(* Logix 5000 project; controller TFF vendor 1 type 14 code 107 rev 33.11; software revision 33.04; part 12 of 38 *)

        [5,197].Criteria2Value := -1000000.0, [5,197].ActionValue := -1000000.0, [5,198].Criteria1 := -999, [5,198].Criteria1Operator := -999, [5,198].Boolean := -999, [5,198].Criteria2 := -999, [5,198].Criteria2Operator := -999, [5,198].Action := -999, [5,198].Label := -999, [5,198].Criteria1Value := -1000000.0, [5,198].Criteria2Value := -1000000.0, [5,198].ActionValue := -1000000.0, [5,199].Criteria1 := -999, [5,199].Criteria1Operator := -999, [5,199].Boolean := -999, [5,199].Criteria2 := -999, [5,199].Criteria2Operator := -999, [5,199].Action := -999, [5,199].Label := -999, [5,199].Criteria1Value := -1000000.0, [5,199].Criteria2Value := -1000000.0, [5,199].ActionValue := -1000000.0, [5,200].Criteria1 := -999, [5,200].Criteria1Operator := -999, [5,200].Boolean := -999, [5,200].Criteria2 := -999, [5,200].Criteria2Operator := -999, [5,200].Action := -999, [5,200].Label := -999, [5,200].Criteria1Value := -1000000.0, [5,200].Criteria2Value := -1000000.0, [5,200].ActionValue := -1000000.0, [5,201].Criteria1 := -999, [5,201].Criteria1Operator := -999, [5,201].Boolean := -999, [5,201].Criteria2 := -999, [5,201].Criteria2Operator := -999, [5,201].Action := -999, [5,201].Label := -999, [5,201].Criteria1Value := -1000000.0, [5,201].Criteria2Value := -1000000.0, [5,201].ActionValue := -1000000.0, [5,202].Criteria1 := -999, [5,202].Criteria1Operator := -999, [5,202].Boolean := -999, [5,202].Criteria2 := -999, [5,202].Criteria2Operator := -999, [5,202].Action := -999, [5,202].Label := -999, [5,202].Criteria1Value := -1000000.0, [5,202].Criteria2Value := -1000000.0, [5,202].ActionValue := -1000000.0, [5,203].Criteria1 := -999, [5,203].Criteria1Operator := -999, [5,203].Boolean := -999, [5,203].Criteria2 := -999, [5,203].Criteria2Operator := -999, [5,203].Action := -999, [5,203].Label := -999, [5,203].Criteria1Value := -1000000.0,
        [5,203].Criteria2Value := -1000000.0, [5,203].ActionValue := -1000000.0, [5,204].Criteria1 := -999, [5,204].Criteria1Operator := -999, [5,204].Boolean := -999, [5,204].Criteria2 := -999, [5,204].Criteria2Operator := -999, [5,204].Action := -999, [5,204].Label := -999, [5,204].Criteria1Value := -1000000.0, [5,204].Criteria2Value := -1000000.0, [5,204].ActionValue := -1000000.0, [5,205].Criteria1 := -999, [5,205].Criteria1Operator := -999, [5,205].Boolean := -999, [5,205].Criteria2 := -999, [5,205].Criteria2Operator := -999, [5,205].Action := -999, [5,205].Label := -999, [5,205].Criteria1Value := -1000000.0, [5,205].Criteria2Value := -1000000.0, [5,205].ActionValue := -1000000.0, [5,206].Criteria1 := -999, [5,206].Criteria1Operator := -999, [5,206].Boolean := -999, [5,206].Criteria2 := -999, [5,206].Criteria2Operator := -999, [5,206].Action := -999, [5,206].Label := -999, [5,206].Criteria1Value := -1000000.0, [5,206].Criteria2Value := -1000000.0, [5,206].ActionValue := -1000000.0, [5,207].Criteria1 := -999, [5,207].Criteria1Operator := -999, [5,207].Boolean := -999, [5,207].Criteria2 := -999, [5,207].Criteria2Operator := -999, [5,207].Action := -999, [5,207].Label := -999, [5,207].Criteria1Value := -1000000.0, [5,207].Criteria2Value := -1000000.0, [5,207].ActionValue := -1000000.0, [5,208].Criteria1 := -999, [5,208].Criteria1Operator := -999, [5,208].Boolean := -999, [5,208].Criteria2 := -999, [5,208].Criteria2Operator := -999, [5,208].Action := -999, [5,208].Label := -999, [5,208].Criteria1Value := -1000000.0, [5,208].Criteria2Value := -1000000.0, [5,208].ActionValue := -1000000.0, [5,209].Criteria1 := -999, [5,209].Criteria1Operator := -999, [5,209].Boolean := -999, [5,209].Criteria2 := -999, [5,209].Criteria2Operator := -999, [5,209].Action := -999, [5,209].Label := -999, [5,209].Criteria1Value := -1000000.0,
        [5,209].Criteria2Value := -1000000.0, [5,209].ActionValue := -1000000.0, [5,210].Criteria1 := -999, [5,210].Criteria1Operator := -999, [5,210].Boolean := -999, [5,210].Criteria2 := -999, [5,210].Criteria2Operator := -999, [5,210].Action := -999, [5,210].Label := -999, [5,210].Criteria1Value := -1000000.0, [5,210].Criteria2Value := -1000000.0, [5,210].ActionValue := -1000000.0, [5,211].Criteria1 := -999, [5,211].Criteria1Operator := -999, [5,211].Boolean := -999, [5,211].Criteria2 := -999, [5,211].Criteria2Operator := -999, [5,211].Action := -999, [5,211].Label := -999, [5,211].Criteria1Value := -1000000.0, [5,211].Criteria2Value := -1000000.0, [5,211].ActionValue := -1000000.0, [5,212].Criteria1 := -999, [5,212].Criteria1Operator := -999, [5,212].Boolean := -999, [5,212].Criteria2 := -999, [5,212].Criteria2Operator := -999, [5,212].Action := -999, [5,212].Label := -999, [5,212].Criteria1Value := -1000000.0, [5,212].Criteria2Value := -1000000.0, [5,212].ActionValue := -1000000.0, [5,213].Criteria1 := -999, [5,213].Criteria1Operator := -999, [5,213].Boolean := -999, [5,213].Criteria2 := -999, [5,213].Criteria2Operator := -999, [5,213].Action := -999, [5,213].Label := -999, [5,213].Criteria1Value := -1000000.0, [5,213].Criteria2Value := -1000000.0, [5,213].ActionValue := -1000000.0, [5,214].Criteria1 := -999, [5,214].Criteria1Operator := -999, [5,214].Boolean := -999, [5,214].Criteria2 := -999, [5,214].Criteria2Operator := -999, [5,214].Action := -999, [5,214].Label := -999, [5,214].Criteria1Value := -1000000.0, [5,214].Criteria2Value := -1000000.0, [5,214].ActionValue := -1000000.0, [5,215].Criteria1 := -999, [5,215].Criteria1Operator := -999, [5,215].Boolean := -999, [5,215].Criteria2 := -999, [5,215].Criteria2Operator := -999, [5,215].Action := -999, [5,215].Label := -999, [5,215].Criteria1Value := -1000000.0,
        [5,215].Criteria2Value := -1000000.0, [5,215].ActionValue := -1000000.0, [5,216].Criteria1 := -999, [5,216].Criteria1Operator := -999, [5,216].Boolean := -999, [5,216].Criteria2 := -999, [5,216].Criteria2Operator := -999, [5,216].Action := -999, [5,216].Label := -999, [5,216].Criteria1Value := -1000000.0, [5,216].Criteria2Value := -1000000.0, [5,216].ActionValue := -1000000.0, [5,217].Criteria1 := -999, [5,217].Criteria1Operator := -999, [5,217].Boolean := -999, [5,217].Criteria2 := -999, [5,217].Criteria2Operator := -999, [5,217].Action := -999, [5,217].Label := -999, [5,217].Criteria1Value := -1000000.0, [5,217].Criteria2Value := -1000000.0, [5,217].ActionValue := -1000000.0, [5,218].Criteria1 := -999, [5,218].Criteria1Operator := -999, [5,218].Boolean := -999, [5,218].Criteria2 := -999, [5,218].Criteria2Operator := -999, [5,218].Action := -999, [5,218].Label := -999, [5,218].Criteria1Value := -1000000.0, [5,218].Criteria2Value := -1000000.0, [5,218].ActionValue := -1000000.0, [5,219].Criteria1 := -999, [5,219].Criteria1Operator := -999, [5,219].Boolean := -999, [5,219].Criteria2 := -999, [5,219].Criteria2Operator := -999, [5,219].Action := -999, [5,219].Label := -999, [5,219].Criteria1Value := -1000000.0, [5,219].Criteria2Value := -1000000.0, [5,219].ActionValue := -1000000.0, [5,220].Criteria1 := -999, [5,220].Criteria1Operator := -999, [5,220].Boolean := -999, [5,220].Criteria2 := -999, [5,220].Criteria2Operator := -999, [5,220].Action := -999, [5,220].Label := -999, [5,220].Criteria1Value := -1000000.0, [5,220].Criteria2Value := -1000000.0, [5,220].ActionValue := -1000000.0, [5,221].Criteria1 := -999, [5,221].Criteria1Operator := -999, [5,221].Boolean := -999, [5,221].Criteria2 := -999, [5,221].Criteria2Operator := -999, [5,221].Action := -999, [5,221].Label := -999, [5,221].Criteria1Value := -1000000.0,
        [5,221].Criteria2Value := -1000000.0, [5,221].ActionValue := -1000000.0, [5,222].Criteria1 := -999, [5,222].Criteria1Operator := -999, [5,222].Boolean := -999, [5,222].Criteria2 := -999, [5,222].Criteria2Operator := -999, [5,222].Action := -999, [5,222].Label := -999, [5,222].Criteria1Value := -1000000.0, [5,222].Criteria2Value := -1000000.0, [5,222].ActionValue := -1000000.0, [5,223].Criteria1 := -999, [5,223].Criteria1Operator := -999, [5,223].Boolean := -999, [5,223].Criteria2 := -999, [5,223].Criteria2Operator := -999, [5,223].Action := -999, [5,223].Label := -999, [5,223].Criteria1Value := -1000000.0, [5,223].Criteria2Value := -1000000.0, [5,223].ActionValue := -1000000.0, [5,224].Criteria1 := -999, [5,224].Criteria1Operator := -999, [5,224].Boolean := -999, [5,224].Criteria2 := -999, [5,224].Criteria2Operator := -999, [5,224].Action := -999, [5,224].Label := -999, [5,224].Criteria1Value := -1000000.0, [5,224].Criteria2Value := -1000000.0, [5,224].ActionValue := -1000000.0, [5,225].Criteria1 := -999, [5,225].Criteria1Operator := -999, [5,225].Boolean := -999, [5,225].Criteria2 := -999, [5,225].Criteria2Operator := -999, [5,225].Action := -999, [5,225].Label := -999, [5,225].Criteria1Value := -1000000.0, [5,225].Criteria2Value := -1000000.0, [5,225].ActionValue := -1000000.0, [5,226].Criteria1 := -999, [5,226].Criteria1Operator := -999, [5,226].Boolean := -999, [5,226].Criteria2 := -999, [5,226].Criteria2Operator := -999, [5,226].Action := -999, [5,226].Label := -999, [5,226].Criteria1Value := -1000000.0, [5,226].Criteria2Value := -1000000.0, [5,226].ActionValue := -1000000.0, [5,227].Criteria1 := -999, [5,227].Criteria1Operator := -999, [5,227].Boolean := -999, [5,227].Criteria2 := -999, [5,227].Criteria2Operator := -999, [5,227].Action := -999, [5,227].Label := -999, [5,227].Criteria1Value := -1000000.0,
        [5,227].Criteria2Value := -1000000.0, [5,227].ActionValue := -1000000.0, [5,228].Criteria1 := -999, [5,228].Criteria1Operator := -999, [5,228].Boolean := -999, [5,228].Criteria2 := -999, [5,228].Criteria2Operator := -999, [5,228].Action := -999, [5,228].Label := -999, [5,228].Criteria1Value := -1000000.0, [5,228].Criteria2Value := -1000000.0, [5,228].ActionValue := -1000000.0, [5,229].Criteria1 := -999, [5,229].Criteria1Operator := -999, [5,229].Boolean := -999, [5,229].Criteria2 := -999, [5,229].Criteria2Operator := -999, [5,229].Action := -999, [5,229].Label := -999, [5,229].Criteria1Value := -1000000.0, [5,229].Criteria2Value := -1000000.0, [5,229].ActionValue := -1000000.0, [5,230].Criteria1 := -999, [5,230].Criteria1Operator := -999, [5,230].Boolean := -999, [5,230].Criteria2 := -999, [5,230].Criteria2Operator := -999, [5,230].Action := -999, [5,230].Label := -999, [5,230].Criteria1Value := -1000000.0, [5,230].Criteria2Value := -1000000.0, [5,230].ActionValue := -1000000.0, [5,231].Criteria1 := -999, [5,231].Criteria1Operator := -999, [5,231].Boolean := -999, [5,231].Criteria2 := -999, [5,231].Criteria2Operator := -999, [5,231].Action := -999, [5,231].Label := -999, [5,231].Criteria1Value := -1000000.0, [5,231].Criteria2Value := -1000000.0, [5,231].ActionValue := -1000000.0, [5,232].Criteria1 := -999, [5,232].Criteria1Operator := -999, [5,232].Boolean := -999, [5,232].Criteria2 := -999, [5,232].Criteria2Operator := -999, [5,232].Action := -999, [5,232].Label := -999, [5,232].Criteria1Value := -1000000.0, [5,232].Criteria2Value := -1000000.0, [5,232].ActionValue := -1000000.0, [5,233].Criteria1 := -999, [5,233].Criteria1Operator := -999, [5,233].Boolean := -999, [5,233].Criteria2 := -999, [5,233].Criteria2Operator := -999, [5,233].Action := -999, [5,233].Label := -999, [5,233].Criteria1Value := -1000000.0,
        [5,233].Criteria2Value := -1000000.0, [5,233].ActionValue := -1000000.0, [5,234].Criteria1 := -999, [5,234].Criteria1Operator := -999, [5,234].Boolean := -999, [5,234].Criteria2 := -999, [5,234].Criteria2Operator := -999, [5,234].Action := -999, [5,234].Label := -999, [5,234].Criteria1Value := -1000000.0, [5,234].Criteria2Value := -1000000.0, [5,234].ActionValue := -1000000.0, [5,235].Criteria1 := -999, [5,235].Criteria1Operator := -999, [5,235].Boolean := -999, [5,235].Criteria2 := -999, [5,235].Criteria2Operator := -999, [5,235].Action := -999, [5,235].Label := -999, [5,235].Criteria1Value := -1000000.0, [5,235].Criteria2Value := -1000000.0, [5,235].ActionValue := -1000000.0, [5,236].Criteria1 := -999, [5,236].Criteria1Operator := -999, [5,236].Boolean := -999, [5,236].Criteria2 := -999, [5,236].Criteria2Operator := -999, [5,236].Action := -999, [5,236].Label := -999, [5,236].Criteria1Value := -1000000.0, [5,236].Criteria2Value := -1000000.0, [5,236].ActionValue := -1000000.0, [5,237].Criteria1 := -999, [5,237].Criteria1Operator := -999, [5,237].Boolean := -999, [5,237].Criteria2 := -999, [5,237].Criteria2Operator := -999, [5,237].Action := -999, [5,237].Label := -999, [5,237].Criteria1Value := -1000000.0, [5,237].Criteria2Value := -1000000.0, [5,237].ActionValue := -1000000.0, [5,238].Criteria1 := -999, [5,238].Criteria1Operator := -999, [5,238].Boolean := -999, [5,238].Criteria2 := -999, [5,238].Criteria2Operator := -999, [5,238].Action := -999, [5,238].Label := -999, [5,238].Criteria1Value := -1000000.0, [5,238].Criteria2Value := -1000000.0, [5,238].ActionValue := -1000000.0, [5,239].Criteria1 := -999, [5,239].Criteria1Operator := -999, [5,239].Boolean := -999, [5,239].Criteria2 := -999, [5,239].Criteria2Operator := -999, [5,239].Action := -999, [5,239].Label := -999, [5,239].Criteria1Value := -1000000.0,
        [5,239].Criteria2Value := -1000000.0, [5,239].ActionValue := -1000000.0, [5,240].Criteria1 := -999, [5,240].Criteria1Operator := -999, [5,240].Boolean := -999, [5,240].Criteria2 := -999, [5,240].Criteria2Operator := -999, [5,240].Action := -999, [5,240].Label := -999, [5,240].Criteria1Value := -1000000.0, [5,240].Criteria2Value := -1000000.0, [5,240].ActionValue := -1000000.0, [5,241].Criteria1 := -999, [5,241].Criteria1Operator := -999, [5,241].Boolean := -999, [5,241].Criteria2 := -999, [5,241].Criteria2Operator := -999, [5,241].Action := -999, [5,241].Label := -999, [5,241].Criteria1Value := -1000000.0, [5,241].Criteria2Value := -1000000.0, [5,241].ActionValue := -1000000.0, [5,242].Criteria1 := -999, [5,242].Criteria1Operator := -999, [5,242].Boolean := -999, [5,242].Criteria2 := -999, [5,242].Criteria2Operator := -999, [5,242].Action := -999, [5,242].Label := -999, [5,242].Criteria1Value := -1000000.0, [5,242].Criteria2Value := -1000000.0, [5,242].ActionValue := -1000000.0, [5,243].Criteria1 := -999, [5,243].Criteria1Operator := -999, [5,243].Boolean := -999, [5,243].Criteria2 := -999, [5,243].Criteria2Operator := -999, [5,243].Action := -999, [5,243].Label := -999, [5,243].Criteria1Value := -1000000.0, [5,243].Criteria2Value := -1000000.0, [5,243].ActionValue := -1000000.0, [5,244].Criteria1 := -999, [5,244].Criteria1Operator := -999, [5,244].Boolean := -999, [5,244].Criteria2 := -999, [5,244].Criteria2Operator := -999, [5,244].Action := -999, [5,244].Label := -999, [5,244].Criteria1Value := -1000000.0, [5,244].Criteria2Value := -1000000.0, [5,244].ActionValue := -1000000.0, [5,245].Criteria1 := -999, [5,245].Criteria1Operator := -999, [5,245].Boolean := -999, [5,245].Criteria2 := -999, [5,245].Criteria2Operator := -999, [5,245].Action := -999, [5,245].Label := -999, [5,245].Criteria1Value := -1000000.0,
        [5,245].Criteria2Value := -1000000.0, [5,245].ActionValue := -1000000.0, [5,246].Criteria1 := -999, [5,246].Criteria1Operator := -999, [5,246].Boolean := -999, [5,246].Criteria2 := -999, [5,246].Criteria2Operator := -999, [5,246].Action := -999, [5,246].Label := -999, [5,246].Criteria1Value := -1000000.0, [5,246].Criteria2Value := -1000000.0, [5,246].ActionValue := -1000000.0, [5,247].Criteria1 := -999, [5,247].Criteria1Operator := -999, [5,247].Boolean := -999, [5,247].Criteria2 := -999, [5,247].Criteria2Operator := -999, [5,247].Action := -999, [5,247].Label := -999, [5,247].Criteria1Value := -1000000.0, [5,247].Criteria2Value := -1000000.0, [5,247].ActionValue := -1000000.0, [5,248].Criteria1 := -999, [5,248].Criteria1Operator := -999, [5,248].Boolean := -999, [5,248].Criteria2 := -999, [5,248].Criteria2Operator := -999, [5,248].Action := -999, [5,248].Label := -999, [5,248].Criteria1Value := -1000000.0, [5,248].Criteria2Value := -1000000.0, [5,248].ActionValue := -1000000.0, [5,249].Criteria1 := -999, [5,249].Criteria1Operator := -999, [5,249].Boolean := -999, [5,249].Criteria2 := -999, [5,249].Criteria2Operator := -999, [5,249].Action := -999, [5,249].Label := -999, [5,249].Criteria1Value := -1000000.0, [5,249].Criteria2Value := -1000000.0, [5,249].ActionValue := -1000000.0, [5,250].Criteria1 := -999, [5,250].Criteria1Operator := -999, [5,250].Boolean := -999, [5,250].Criteria2 := -999, [5,250].Criteria2Operator := -999, [5,250].Action := -999, [5,250].Label := -999, [5,250].Criteria1Value := -1000000.0, [5,250].Criteria2Value := -1000000.0, [5,250].ActionValue := -1000000.0);   // Operation Table
        [0,0]   // Null Step
        [1,0]   // Null Step
        [2,0]   // Null Step
        [3,0]   // Null Step
        [4,0]   // Null Step
        [5,0]   // Null Step
   Options : Options := (CCP_Report := 1, InletFeed := 1, FeedTank := 1, TransferFlow := 1, TankPH := 1, FiltrateNoInstrum_Dis := 1, FiltrateCondPHUV := 1, FiltrateUltrasonicFlow := 1, SingleUsePH := 1, External_IO := 1, TFF80 := 1);   // Options List
   PCDateTime : DINT[7] := ([0] := 2025, [1] := 10, [2] := 3, [3] := 11, [4] := 41, [5] := 1, [6] := -1);   // Date/Time Array from PC
   PcToPLCHeartBeat : BOOL;   // PC to PLC communication heartbeat Set to 1 by HMI Reset to 0 by plc
   PCV101 : ALIAS FOR AnalogPoint[3];
   PCV101_AO : ALIAS FOR AnalogOutput[3];
   PCV101_Calib : PCV_Calib;   // PCV101 Position Calibration
   PCV101_Control : PCV_Control := (FullOpenResetTimer.PRE := 3000, FullCloseSP := 100.0, FullCloseResetTimer.PRE := 3000, ClosedStatusSP := 95.0);   // PCV101 Control UDT
   PCV101_CVTune : CVTune := (ClosedRaw := 12340.0, OpenRaw := 27508.0, MaxOutput := 100.0, MinTimer.PRE := 5000, MaxTimer.PRE := 5000);
   PCV101_PID : PCV := (PV := 0.032964136, CV := 100.0, OpenRawValue := 27508.0, ClosedRawValue := 12340.0);   // PCV101 PID Management
   PCV101_SIG : ALIAS FOR DigitalPoint[102];
   PCV101Alarm : ALIAS FOR AlarmAnalog[3];
   PCV201 : ALIAS FOR AnalogPoint[4];
   PCV201_AO : ALIAS FOR AnalogOutput[4];
   PCV201_Calib : PCV_Calib;   // PCV201 Position Calibration
   PCV201_Control : PCV_Control := (FullOpenSP := 100.0, FullOpenResetTimer.PRE := 3000, FullCloseResetTimer.PRE := 3000, ClosedStatusSP := 95.0);   // PCV201 Control UDT
   PCV201_CVTune : CVTune := (ClosedRaw := 25520.0, OpenRaw := 10318.0, MaxOutput := 100.0, MinTimer.PRE := 5000, MaxTimer.PRE := 5000);
   PCV201_PID : PCV := (PV := 51.769505, OpenRawValue := 10318.0, ClosedRawValue := 25520.0);   // PCV201 PID Management
   PCV201_SIG : ALIAS FOR DigitalPoint[103];
   PCV201Alarm : ALIAS FOR AlarmAnalog[4];
   PERM : ALIAS FOR AnalogPoint[46];
   PERMAlarm : ALIAS FOR AlarmAnalog[46];
   Phase : Phases[6] := ([0].Stop := 1, [0].Hold := 1, [0].JumpStep := 13, [0].StartStep := 1, [0].TotalSteps := 16, [0].ActualStep := 12, [1].JumpStep := 51, [1].StartStep := 1, [1].TotalSteps := 49, [1].ActualStep := 50, [2].JumpStep := 11, [2].StartStep := 1, [2].TotalSteps := 9, [2].ActualStep := 10, [3].JumpStep := 14, [3].StartStep := 1, [3].TotalSteps := 45, [3].ActualStep := 13, [4].JumpStep := 68, [4].StartStep := 1, [4].TotalSteps := 66, [4].ActualStep := 67, [5].JumpStep := 6, [5].StartStep := 1, [5].Crit1MetTime := 1, [5].ActualStep := 5);   // Phase Control Array
   Phase0 : ALIAS FOR Phase[0];   // Phase 0
   Phase0_PauseTime : ALIAS FOR Timers[12];   // Phase 0 Pause Time
   Phase0_StepTime : ALIAS FOR Timers[6];   // Phase 0 Step Time
   Phase0_Totalizer_Feed : ALIAS FOR PhaseTotalizer[0];   // Phase 0 Total Feed
   Phase0_Totalizer_Filtrate : ALIAS FOR PhaseTotalizer[6];   // Phase 0 Total Filtrate
   Phase0_Totalizer_Transfer : ALIAS FOR PhaseTotalizer[12];   // Phase 0 Total Transfer
   Phase0_TotalTime : ALIAS FOR Timers[0];   // Phase 0 Total Time
   Phase1 : ALIAS FOR Phase[1];   // Phase 1
   Phase1_PauseTime : ALIAS FOR Timers[13];   // Phase 1 Pause Time
   Phase1_StepTime : ALIAS FOR Timers[7];   // Phase 1 Step Time
   Phase1_Totalizer_Feed : ALIAS FOR PhaseTotalizer[1];   // Phase 1 Total Feed
   Phase1_Totalizer_Filtrate : ALIAS FOR PhaseTotalizer[7];   // Phase 1 Total Filtrate
   Phase1_Totalizer_Transfer : ALIAS FOR PhaseTotalizer[13];   // Phase 1 Total Transfer
   Phase1_TotalTime : ALIAS FOR Timers[1];   // Phase 1 Total Time
   Phase2 : ALIAS FOR Phase[2];   // Phase 2
   Phase2_PauseTime : ALIAS FOR Timers[14];   // Phase 2 Pause Time
   Phase2_StepTime : ALIAS FOR Timers[8];   // Phase 2 Step Time
   Phase2_Totalizer_Feed : ALIAS FOR PhaseTotalizer[2];   // Phase 2 Total Feed
   Phase2_Totalizer_Filtrate : ALIAS FOR PhaseTotalizer[8];   // Phase 2 Total Filtrate
   Phase2_Totalizer_Transfer : ALIAS FOR PhaseTotalizer[14];   // Phase 2 Total Transfer
   Phase2_TotalTime : ALIAS FOR Timers[2];   // Phase 2 Total Time
   Phase3 : ALIAS FOR Phase[3];   // Phase 3
   Phase3_PauseTime : ALIAS FOR Timers[15];   // Phase 3 Pause Time
   Phase3_StepTime : ALIAS FOR Timers[9];   // Phase 3 Step Time
   Phase3_Totalizer_Feed : ALIAS FOR PhaseTotalizer[3];   // Phase 3 Total Feed
   Phase3_Totalizer_Filtrate : ALIAS FOR PhaseTotalizer[9];   // Phase 3 Total Filtrate
   Phase3_Totalizer_Transfer : ALIAS FOR PhaseTotalizer[15];   // Phase 3 Total Transfer
   Phase3_TotalTime : ALIAS FOR Timers[3];   // Phase 3 Total Time
   Phase4 : ALIAS FOR Phase[4];   // Phase 4
   Phase4_PauseTime : ALIAS FOR Timers[16];   // Phase 4 Pause Time
   Phase4_StepTime : ALIAS FOR Timers[10];   // Phase 4 Step Time
   Phase4_Totalizer_Feed : ALIAS FOR PhaseTotalizer[4];   // Phase 4 Total Feed
   Phase4_Totalizer_Filtrate : ALIAS FOR PhaseTotalizer[10];   // Phase 4 Total Filtrate
   Phase4_Totalizer_Transfer : ALIAS FOR PhaseTotalizer[16];   // Phase 4 Total Transfer
   Phase4_TotalTime : ALIAS FOR Timers[4];   // Phase 4 Total Time
   Phase5 : ALIAS FOR Phase[5];   // Phase 5
   Phase5_PauseTime : ALIAS FOR Timers[17];   // Phase 5 Pause Time
   Phase5_StepTime : ALIAS FOR Timers[11];   // Phase 5 Step Time
   Phase5_Totalizer_Feed : ALIAS FOR PhaseTotalizer[5];   // Phase 5 Total Feed
   Phase5_Totalizer_Filtrate : ALIAS FOR PhaseTotalizer[11];   // Phase 5 Total Filtrate
   Phase5_Totalizer_Transfer : ALIAS FOR PhaseTotalizer[17];   // Phase 5 Total Transfer
   Phase5_TotalTime : ALIAS FOR Timers[5];   // Phase 5 Total Time
   PhaseTotalizer : PhaseTotalizer[18] := ([0].Enable := 1, [0].PVscale := 60.0, [0].Title := 'Phase0 Vol', [0].EGU := 'L', [0].EnableCfg := 1, [0].SourceAddressCfg := 42, [1].Enable := 1, [1].PVscale := 60.0, [1].Title := 'Phase1 Vol', [1].EGU := 'L', [1].EnableCfg := 1, [1].SourceAddressCfg := 42, [2].PVscale := 60.0, [2].Title := 'Phase2 Vol', [2].EGU := 'L', [2].EnableCfg := 1, [2].SourceAddressCfg := 42, [3].PVscale := 60.0, [3].Title := 'Phase3 Vol', [3].EGU := 'L', [3].EnableCfg := 1, [3].SourceAddressCfg := 42, [4].PVscale := 60.0, [4].Title := 'Phase4 Vol', [4].EGU := 'L', [4].EnableCfg := 1, [4].SourceAddressCfg := 42, [5].PVscale := 60.0, [5].Title := 'Phase5 Vol', [5].EGU := 'L', [5].EnableCfg := 1, [5].SourceAddressCfg := 42, [6].Enable := 1, [6].PV := -23.77737, [6].PVscale := 60.0, [6].Title := 'Phase0 Vol', [6].EGU := 'L', [6].EnableCfg := 1, [6].SourceAddressCfg := 2, [7].PV := -23.77737, [7].PVscale := 60.0, [7].Title := 'Phase1 Vol', [7].EGU := 'L', [7].EnableCfg := 1, [7].SourceAddressCfg := 2, [8].PV := -23.77737, [8].PVscale := 60.0, [8].Title := 'Phase2 Vol', [8].EGU := 'L', [8].EnableCfg := 1, [8].SourceAddressCfg := 2, [9].PV := -23.77737, [9].PVscale := 60.0, [9].Title := 'Phase3 Vol', [9].EGU := 'L', [9].EnableCfg := 1, [9].SourceAddressCfg := 2, [10].PV := -23.77737, [10].PVscale := 60.0, [10].Title := 'Phase4 Vol',
        [10].EGU := 'L', [10].EnableCfg := 1, [10].SourceAddressCfg := 2, [11].PV := -23.77737, [11].PVscale := 60.0, [11].Title := 'Phase5 Vol', [11].EGU := 'L', [11].EnableCfg := 1, [11].SourceAddressCfg := 2, [12].PVscale := 60.0, [12].EnableCfg := 1, [12].SourceAddressCfg := 20, [13].PVscale := 60.0, [13].EnableCfg := 1, [13].SourceAddressCfg := 20, [14].PVscale := 60.0, [14].EnableCfg := 1, [14].SourceAddressCfg := 20, [15].PVscale := 60.0, [15].EnableCfg := 1, [15].SourceAddressCfg := 20, [16].PVscale := 60.0, [16].EnableCfg := 1, [16].SourceAddressCfg := 20, [17].PVscale := 60.0, [17].EnableCfg := 1, [17].SourceAddressCfg := 20);   // Phase Totalizers Array
        [0]   // Phase 0 Totalizer 1
        [1]   // Phase 1 Totalizer 1
        [10]   // Phase 4 Totalizer 2
        [11]   // Phase 5 Totalizer 2
        [12]   // Phase 0 Totalizer 3
        [13]   // Phase 1 Totalizer 3
        [14]   // Phase 2 Totalizer 3
        [2]   // Phase 2 Totalizer 1
        [3]   // Phase 3 Totalizer 1
        [4]   // Phase 4 Totalizer 1
        [5]   // Phase 5 Totalizer 1
        [6]   // Phase 0 Totalizer 2
        [7]   // Phase 1 Totalizer 2
        [8]   // Phase 2 Totalizer 2
        [9]   // Phase 3 Totalizer 2
        [15]   // Phase 3 Totalizer 3
        [16]   // Phase 4 Totalizer 3
        [17]   // Phase 5 Totalizer 3
   PhaseTotalizer_Storage : PhaseTotalizer[6,18] := ([0,0].Enable := 1, [0,0].PVscale := 60.0, [0,0].Title := 'Phase0 Vol', [0,0].EGU := 'L', [0,0].EnableCfg := 1, [0,0].SourceAddressCfg := 40, [0,1].Enable := 1, [0,1].PVscale := 60.0, [0,1].Title := 'Phase1 Vol', [0,1].EGU := 'L', [0,1].EnableCfg := 1, [0,1].SourceAddressCfg := 40, [0,2].PVscale := 60.0, [0,2].Title := 'Phase2 Vol', [0,2].EGU := 'L', [0,2].EnableCfg := 1, [0,2].SourceAddressCfg := 40, [0,3].PVscale := 60.0, [0,3].Title := 'Phase3 Vol', [0,3].EGU := 'L', [0,3].EnableCfg := 1, [0,3].SourceAddressCfg := 40, [0,4].PVscale := 60.0, [0,4].Title := 'Phase4 Vol', [0,4].EGU := 'L', [0,4].EnableCfg := 1, [0,4].SourceAddressCfg := 40, [0,5].PVscale := 60.0, [0,5].Title := 'Phase5 Vol', [0,5].EGU := 'L', [0,5].EnableCfg := 1, [0,5].SourceAddressCfg := 40, [0,6].Enable := 1, [0,6].PVscale := 60.0, [0,6].Title := 'Phase0 CVs', [0,6].EGU := 'CVs', [0,6].EnableCfg := 1, [0,6].SourceTypeCfg := 1, [0,7].PVscale := 60.0, [0,7].Title := 'Phase1 CVs', [0,7].EGU := 'CVs', [0,7].EnableCfg := 1, [0,7].SourceTypeCfg := 1, [0,8].PVscale := 60.0, [0,8].Title := 'Phase2 CVs', [0,8].EGU := 'CVs', [0,8].EnableCfg := 1, [0,8].SourceTypeCfg := 1, [0,9].PVscale := 60.0, [0,9].Title := 'Phase3 CVs', [0,9].EGU := 'CVs', [0,9].EnableCfg := 1, [0,9].SourceTypeCfg := 1, [0,10].PVscale := 60.0, [0,10].Title := 'Phase4 CVs', [0,10].EGU := 'CVs', [0,10].EnableCfg := 1, [0,10].SourceTypeCfg := 1, [0,11].PVscale := 60.0, [0,11].Title := 'Phase5 CVs',
        [0,11].EGU := 'CVs', [0,11].EnableCfg := 1, [0,11].SourceTypeCfg := 1, [1,0].Enable := 1, [1,0].PVscale := 60.0, [1,0].Title := 'Phase0 Vol', [1,0].EGU := 'L', [1,0].EnableCfg := 1, [1,0].SourceAddressCfg := 40, [1,1].Enable := 1, [1,1].PVscale := 60.0, [1,1].Title := 'Phase1 Vol', [1,1].EGU := 'L', [1,1].EnableCfg := 1, [1,1].SourceAddressCfg := 40, [1,2].PVscale := 60.0, [1,2].Title := 'Phase2 Vol', [1,2].EGU := 'L', [1,2].EnableCfg := 1, [1,2].SourceAddressCfg := 40, [1,3].PVscale := 60.0, [1,3].Title := 'Phase3 Vol', [1,3].EGU := 'L', [1,3].EnableCfg := 1, [1,3].SourceAddressCfg := 40, [1,4].PVscale := 60.0, [1,4].Title := 'Phase4 Vol', [1,4].EGU := 'L', [1,4].EnableCfg := 1, [1,4].SourceAddressCfg := 40, [1,5].PVscale := 60.0, [1,5].Title := 'Phase5 Vol', [1,5].EGU := 'L', [1,5].EnableCfg := 1, [1,5].SourceAddressCfg := 40, [1,6].Enable := 1, [1,6].PVscale := 60.0, [1,6].Title := 'Phase0 CVs', [1,6].EGU := 'CVs', [1,6].EnableCfg := 1, [1,6].SourceTypeCfg := 1, [1,7].PVscale := 60.0, [1,7].Title := 'Phase1 CVs', [1,7].EGU := 'CVs', [1,7].EnableCfg := 1, [1,7].SourceTypeCfg := 1, [1,8].PVscale := 60.0, [1,8].Title := 'Phase2 CVs', [1,8].EGU := 'CVs', [1,8].EnableCfg := 1, [1,8].SourceTypeCfg := 1, [1,9].PVscale := 60.0, [1,9].Title := 'Phase3 CVs', [1,9].EGU := 'CVs', [1,9].EnableCfg := 1, [1,9].SourceTypeCfg := 1, [1,10].PVscale := 60.0, [1,10].Title := 'Phase4 CVs', [1,10].EGU := 'CVs', [1,10].EnableCfg := 1,
        [1,10].SourceTypeCfg := 1, [1,11].PVscale := 60.0, [1,11].Title := 'Phase5 CVs', [1,11].EGU := 'CVs', [1,11].EnableCfg := 1, [1,11].SourceTypeCfg := 1, [2,0].Enable := 1, [2,0].PVscale := 60.0, [2,0].Title := 'Phase0 Vol', [2,0].EGU := 'L', [2,0].EnableCfg := 1, [2,0].SourceAddressCfg := 40, [2,1].Enable := 1, [2,1].PVscale := 60.0, [2,1].Title := 'Phase1 Vol', [2,1].EGU := 'L', [2,1].EnableCfg := 1, [2,1].SourceAddressCfg := 40, [2,2].PVscale := 60.0, [2,2].Title := 'Phase2 Vol', [2,2].EGU := 'L', [2,2].EnableCfg := 1, [2,2].SourceAddressCfg := 40, [2,3].PVscale := 60.0, [2,3].Title := 'Phase3 Vol', [2,3].EGU := 'L', [2,3].EnableCfg := 1, [2,3].SourceAddressCfg := 40, [2,4].PVscale := 60.0, [2,4].Title := 'Phase4 Vol', [2,4].EGU := 'L', [2,4].EnableCfg := 1, [2,4].SourceAddressCfg := 40, [2,5].PVscale := 60.0, [2,5].Title := 'Phase5 Vol', [2,5].EGU := 'L', [2,5].EnableCfg := 1, [2,5].SourceAddressCfg := 40, [2,6].Enable := 1, [2,6].PVscale := 60.0, [2,6].Title := 'Phase0 CVs', [2,6].EGU := 'CVs', [2,6].EnableCfg := 1, [2,6].SourceTypeCfg := 1, [2,7].PVscale := 60.0, [2,7].Title := 'Phase1 CVs', [2,7].EGU := 'CVs', [2,7].EnableCfg := 1, [2,7].SourceTypeCfg := 1, [2,8].PVscale := 60.0, [2,8].Title := 'Phase2 CVs', [2,8].EGU := 'CVs', [2,8].EnableCfg := 1, [2,8].SourceTypeCfg := 1, [2,9].PVscale := 60.0, [2,9].Title := 'Phase3 CVs', [2,9].EGU := 'CVs', [2,9].EnableCfg := 1, [2,9].SourceTypeCfg := 1, [2,10].PVscale := 60.0,
        [2,10].Title := 'Phase4 CVs', [2,10].EGU := 'CVs', [2,10].EnableCfg := 1, [2,10].SourceTypeCfg := 1, [2,11].PVscale := 60.0, [2,11].Title := 'Phase5 CVs', [2,11].EGU := 'CVs', [2,11].EnableCfg := 1, [2,11].SourceTypeCfg := 1, [3,0].PV := 48.590927, [3,0].PVscale := 60.0, [3,0].PVsec := 0.8098488, [3,0].EnableCfg := 1, [3,0].SourceAddressCfg := 40, [3,1].PV := 48.590927, [3,1].PVscale := 60.0, [3,1].PVsec := 0.8098488, [3,1].EnableCfg := 1, [3,1].SourceAddressCfg := 40, [3,2].PV := 48.590927, [3,2].PVscale := 60.0, [3,2].PVsec := 0.8098488, [3,2].EnableCfg := 1, [3,2].SourceAddressCfg := 40, [3,3].PV := 48.590927, [3,3].PVscale := 60.0, [3,3].PVsec := 0.8098488, [3,3].EnableCfg := 1, [3,3].SourceAddressCfg := 40, [3,4].PV := 48.590927, [3,4].PVscale := 60.0, [3,4].PVsec := 0.8098488, [3,4].EnableCfg := 1, [3,4].SourceAddressCfg := 40, [3,5].PV := 48.590927, [3,5].PVscale := 60.0, [3,5].PVsec := 0.8098488, [3,5].EnableCfg := 1, [3,5].SourceAddressCfg := 40, [3,6].PV := 4.8590927, [3,6].PVscale := 60.0, [3,6].PVsec := 0.080984876, [3,6].EnableCfg := 1, [3,6].SourceTypeCfg := 1, [3,7].PV := 4.8590927, [3,7].PVscale := 60.0, [3,7].PVsec := 0.080984876, [3,7].EnableCfg := 1, [3,7].SourceTypeCfg := 1, [3,8].PV := 4.8590927, [3,8].PVscale := 60.0, [3,8].PVsec := 0.080984876, [3,8].EnableCfg := 1, [3,8].SourceTypeCfg := 1, [3,9].PV := 4.8590927, [3,9].PVscale := 60.0, [3,9].PVsec := 0.080984876, [3,9].EnableCfg := 1, [3,9].SourceTypeCfg := 1, [3,10].PV := 4.8590927,
        [3,10].PVscale := 60.0, [3,10].PVsec := 0.080984876, [3,10].EnableCfg := 1, [3,10].SourceTypeCfg := 1, [3,11].PV := 4.8590927, [3,11].PVscale := 60.0, [3,11].PVsec := 0.080984876, [3,11].EnableCfg := 1, [3,11].SourceTypeCfg := 1, [4,0].Enable := 1, [4,0].PVscale := 60.0, [4,0].Title := 'Phase0 Vol', [4,0].EGU := 'L', [4,0].EnableCfg := 1, [4,0].SourceAddressCfg := 40, [4,1].Enable := 1, [4,1].PVscale := 60.0, [4,1].Title := 'Phase1 Vol', [4,1].EGU := 'L', [4,1].EnableCfg := 1, [4,1].SourceAddressCfg := 40, [4,2].PVscale := 60.0, [4,2].Title := 'Phase2 Vol', [4,2].EGU := 'L', [4,2].EnableCfg := 1, [4,2].SourceAddressCfg := 40, [4,3].PVscale := 60.0, [4,3].Title := 'Phase3 Vol', [4,3].EGU := 'L', [4,3].EnableCfg := 1, [4,3].SourceAddressCfg := 40, [4,4].PVscale := 60.0, [4,4].Title := 'Phase4 Vol', [4,4].EGU := 'L', [4,4].EnableCfg := 1, [4,4].SourceAddressCfg := 40, [4,5].PVscale := 60.0, [4,5].Title := 'Phase5 Vol', [4,5].EGU := 'L', [4,5].EnableCfg := 1, [4,5].SourceAddressCfg := 40, [4,6].Enable := 1, [4,6].PVscale := 60.0, [4,6].Title := 'Phase0 CVs', [4,6].EGU := 'CVs', [4,6].EnableCfg := 1, [4,6].SourceTypeCfg := 1, [4,7].PVscale := 60.0, [4,7].Title := 'Phase1 CVs', [4,7].EGU := 'CVs', [4,7].EnableCfg := 1, [4,7].SourceTypeCfg := 1, [4,8].PVscale := 60.0, [4,8].Title := 'Phase2 CVs', [4,8].EGU := 'CVs', [4,8].EnableCfg := 1, [4,8].SourceTypeCfg := 1, [4,9].PVscale := 60.0, [4,9].Title := 'Phase3 CVs', [4,9].EGU := 'CVs',
        [4,9].EnableCfg := 1, [4,9].SourceTypeCfg := 1, [4,10].PVscale := 60.0, [4,10].Title := 'Phase4 CVs', [4,10].EGU := 'CVs', [4,10].EnableCfg := 1, [4,10].SourceTypeCfg := 1, [4,11].PVscale := 60.0, [4,11].Title := 'Phase5 CVs', [4,11].EGU := 'CVs', [4,11].EnableCfg := 1, [4,11].SourceTypeCfg := 1, [5,0].Enable := 1, [5,0].PVscale := 60.0, [5,0].Title := 'Phase0 Vol', [5,0].EGU := 'L', [5,0].EnableCfg := 1, [5,0].SourceAddressCfg := 40, [5,1].Enable := 1, [5,1].PVscale := 60.0, [5,1].Title := 'Phase1 Vol', [5,1].EGU := 'L', [5,1].EnableCfg := 1, [5,1].SourceAddressCfg := 40, [5,2].PVscale := 60.0, [5,2].Title := 'Phase2 Vol', [5,2].EGU := 'L', [5,2].EnableCfg := 1, [5,2].SourceAddressCfg := 40, [5,3].PVscale := 60.0, [5,3].Title := 'Phase3 Vol', [5,3].EGU := 'L', [5,3].EnableCfg := 1, [5,3].SourceAddressCfg := 40, [5,4].PVscale := 60.0, [5,4].Title := 'Phase4 Vol', [5,4].EGU := 'L', [5,4].EnableCfg := 1, [5,4].SourceAddressCfg := 40, [5,5].PVscale := 60.0, [5,5].Title := 'Phase5 Vol', [5,5].EGU := 'L', [5,5].EnableCfg := 1, [5,5].SourceAddressCfg := 40, [5,6].Enable := 1, [5,6].PVscale := 60.0, [5,6].Title := 'Phase0 CVs', [5,6].EGU := 'CVs', [5,6].EnableCfg := 1, [5,6].SourceTypeCfg := 1, [5,7].PVscale := 60.0, [5,7].Title := 'Phase1 CVs', [5,7].EGU := 'CVs', [5,7].EnableCfg := 1, [5,7].SourceTypeCfg := 1, [5,8].PVscale := 60.0, [5,8].Title := 'Phase2 CVs', [5,8].EGU := 'CVs', [5,8].EnableCfg := 1, [5,8].SourceTypeCfg := 1,
        [5,9].PVscale := 60.0, [5,9].Title := 'Phase3 CVs', [5,9].EGU := 'CVs', [5,9].EnableCfg := 1, [5,9].SourceTypeCfg := 1, [5,10].PVscale := 60.0, [5,10].Title := 'Phase4 CVs', [5,10].EGU := 'CVs', [5,10].EnableCfg := 1, [5,10].SourceTypeCfg := 1, [5,11].PVscale := 60.0, [5,11].Title := 'Phase5 CVs', [5,11].EGU := 'CVs', [5,11].EnableCfg := 1, [5,11].SourceTypeCfg := 1);
   PI001 : ALIAS FOR AnalogPoint[5];
   PI001_SIG : ALIAS FOR DigitalPoint[97];
   PI001Alarm : ALIAS FOR AlarmAnalog[5];
   PI101 : ALIAS FOR AnalogPoint[6];
   PI101_SIG : ALIAS FOR DigitalPoint[98];
   PI101Alarm : ALIAS FOR AlarmAnalog[6];
   PI201 : ALIAS FOR AnalogPoint[7];
   PI201_SIG : ALIAS FOR DigitalPoint[99];
   PI201Alarm : ALIAS FOR AlarmAnalog[7];
   PI401 : ALIAS FOR AnalogPoint[8];
   PI401_SIG : ALIAS FOR DigitalPoint[100];
   PI401Alarm : ALIAS FOR AlarmAnalog[8];
   PI601 : ALIAS FOR AnalogPoint[21];
   PI601_SIG : ALIAS FOR DigitalPoint[95];
   PI601Alarm : ALIAS FOR AlarmAnalog[21];
   PipeAnimation : PipeAnimation;   // HMI Pipe Animation Array
   PipeStatValueHMI : INT[224];   // Pipe Animation Value For HMI
   PISL601 : ALIAS FOR DigitalPoint[0];
   PISL602 : ALIAS FOR DigitalPoint[1];
   PLCFault : FaultRecordType := (Info[0] := 2, Info[1] := 7162, Info[2] := 26809, Info[3] := 931612);   // PLC Major Fault Record
        .Code   // Unique code for the fault
        .TimeLow   // Lower 32 bits of the fault timestamp value
        .TimeHigh   // Upper 32 bits of the fault timestamp value
        .RecType   // Fault Type
        .Info   // Fault specific information
   POWERON : ALIAS FOR DigitalOutput[1];
   ProcedureTime : ALIAS FOR Timers[19];   // Procedure Time
   Prompt : Prompt[7] := ([3].Flag := 1, [3].Step := 12, [3].Value := 1, [5].Value := 1, [6].Step := 5);   // Prompt Array
   Prompt0 : ALIAS FOR Prompt[0];   // Phase 0 Prompt
   Prompt1 : ALIAS FOR Prompt[1];   // Phase 1 Prompt
   Prompt2 : ALIAS FOR Prompt[2];   // Phase 2 Prompt
   Prompt3 : ALIAS FOR Prompt[3];   // Phase 3 Prompt
   Prompt4 : ALIAS FOR Prompt[4];   // Phase 4 Prompt
   Prompt5 : ALIAS FOR Prompt[5];   // Phase 5 Prompt
   PromptTimer : FBD_TIMER := (PRE := 1000, EN := 1);   // Prompt Timer
   PSH001 : ALIAS FOR DigitalPoint[21];
   PSH401 : ALIAS FOR DigitalPoint[22];
   PTA001 : ALIAS FOR DigitalOutput[21];
   PTA101 : ALIAS FOR DigitalOutput[22];
   PTA201 : ALIAS FOR DigitalOutput[23];
   PTA401 : ALIAS FOR DigitalOutput[24];
   PTA601 : ALIAS FOR DigitalOutput[26];
   PumpRunStatus : DINT;   // Pumps Run Status (1 = At least one pump running , 0 = no pump running)
   Rack_ACT350_WI101_200L : IO_Station := (Node_Comm_Status_value := 12288);   // Status of ACT350 200L
   Rack_ACT350_WI101_500L : IO_Station := (Node_Comm_Status_value := 12288);   // Status of ACT350 500L
   Rack_Murr_Node0_Smart : IO_Station := (Node_Comm_Status_value := 16384, Node_Comm_Status := 1, Node_Internal_Defect_Status_value := -125, MOM_Status := 127, MOM_Enable_Config := 1);   // Status of Node 0 Smart
   Rack_Murr_Node1_TFF : IO_Station := (MOM_Status := 1);   // Node 1 data for MOM Config
   Rack_Murr_Node1_TFF20 : IO_Station := (Node_Comm_Status_value := 12288, Node_Internal_Defect_Status := 1);   // Status of Node 1 TFF20
   Rack_Murr_Node1_TFF40 : IO_Station := (Node_Comm_Status_value := 12288, Node_Internal_Defect_Status := 1);   // Status of Node 1 TFF40
   Rack_Murr_Node1_TFF80 : IO_Station := (Node_Comm_Status_value := 16384, Node_Comm_Status := 1, Node_Internal_Defect_Status_value := 126);   // Status of Node 1 TFF80
   RawAnalogInputArray : INT[50] := ([2] := 320, [3] := 12354, [4] := 17653, [5] := 32767, [6] := 6577, [7] := 6567, [8] := 6563, [19] := 6555, [20] := 6549, [37] := 6414);   // Array of analog input raw
   RecipeStepLog_DateTime : STRING25;
   ResumeDownloadFromHOLD : BOOL;   // Resume Download From HOLD
   RSBUZZ : ALIAS FOR DigitalPoint[3];
   ScaleFiltering : ScaleFiltering := (CurrentFilter := 2, Sample_Rate := 10, Timer.PRE := 99999999, Timer.ACC := 5, Timer.EN := 1, Timer.TT := 1, WI101_Unfiltered := -127.832535, FeedBagVolume := -126.566864, FeedBagVolume_Array[0] := -126.566864, FeedBagVolume_Array[1] := -126.566864, FeedBagVolume_Array[2] := -126.566864, FeedBagVolume_Array[3] := -126.566864, FeedBagVolume_Array[4] := -126.566864, FeedBagVolume_Array[5] := -126.566864, FeedBagVolume_Array[6] := -126.566864, FeedBagVolume_Array[7] := -126.566864, FeedBagVolume_Array[8] := -126.566864, FeedBagVolume_Array[9] := -126.566864, FeedBagVolume_Array[10] := -126.566864, FeedBagVolume_Array[11] := -126.566864, FeedBagVolume_Array[12] := -126.566864, FeedBagVolume_Array[13] := -126.566864, FeedBagVolume_Array[14] := -126.566864, FeedBagVolume_Array[15] := -126.566864, FeedBagVolume_Array[16] := -126.566864, FeedBagVolume_Array[17] := -126.566864, FeedBagVolume_Array[18] := -126.566864, FeedBagVolume_Array[19] := -126.566864, FeedBagVolume_Array[20] := -126.566864, FeedBagVolume_Array[21] := -126.566864, FeedBagVolume_Array[22] := -126.566864, FeedBagVolume_Array[23] := -126.566864, FeedBagVolume_Array[24] := -126.566864, FeedBagVolume_Array[25] := -126.566864, FeedBagVolume_Array[26] := -126.566864, FeedBagVolume_Array[27] := -126.566864, FeedBagVolume_Array[28] := -126.566864, FeedBagVolume_Array[29] := -126.566864, FeedBagVolume_Array[30] := -126.566864, FeedBagVolume_Array[31] := -126.566864, FeedBagVolume_Array[32] := -126.566864, FeedBagVolume_Array[33] := -126.566864, FeedBagVolume_Array[34] := -126.566864, FeedBagVolume_Array[35] := -126.566864, FeedBagVolume_Array[36] := -126.566864, FeedBagVolume_Array[37] := -126.566864, FeedBagVolume_Array[38] := -126.566864, FeedBagVolume_Array[39] := -126.566864, FeedBagVolume_Array[40] := -126.566864, FeedBagVolume_Array[41] := -126.566864, FeedBagVolume_Array[42] := -126.566864, FeedBagVolume_Array[43] := -126.566864, FeedBagVolume_Array[44] := -126.566864, FeedBagVolume_Array[45] := -126.566864, FeedBagVolume_Array[46] := -126.566864, FeedBagVolume_Array[47] := -126.566864, FeedBagVolume_Array[48] := -126.566864, FeedBagVolume_Array[49] := -126.566864, FeedBagVolume_Array[50] := -126.566864, FeedBagVolume_Array[51] := -126.566864,
        FeedBagVolume_Array[52] := -126.566864, FeedBagVolume_Array[53] := -126.566864, FeedBagVolume_Array[54] := -126.566864, FeedBagVolume_Array[55] := -126.566864, FeedBagVolume_Array[56] := -126.566864, FeedBagVolume_Array[57] := -126.566864, FeedBagVolume_Array[58] := -126.566864, FeedBagVolume_Array[59] := -126.566864, FeedBagVolume_Array[60] := -126.566864, FeedBagVolume_Array[61] := -126.566864, FeedBagVolume_Array[62] := -126.566864, FeedBagVolume_Array[63] := -126.566864, FeedBagVolume_Array[64] := -126.566864, FeedBagVolume_Array[65] := -126.566864, FeedBagVolume_Array[66] := -126.566864, FeedBagVolume_Array[67] := -126.566864, FeedBagVolume_Array[68] := -126.566864, FeedBagVolume_Array[69] := -126.566864, FeedBagVolume_Array[70] := -126.566864, FeedBagVolume_Array[71] := -126.566864, FeedBagVolume_Array[72] := -126.566864, FeedBagVolume_Array[73] := -126.566864, FeedBagVolume_Array[74] := -126.566864, FeedBagVolume_Array[75] := -126.566864, FeedBagVolume_Array[76] := -126.566864, FeedBagVolume_Array[77] := -126.566864, FeedBagVolume_Array[78] := -126.566864, FeedBagVolume_Array[79] := -126.566864, FeedBagVolume_Array[80] := -126.566864, FeedBagVolume_Array[81] := -126.566864, FeedBagVolume_Array[82] := -126.566864, FeedBagVolume_Array[83] := -126.566864, FeedBagVolume_Array[84] := -126.566864, FeedBagVolume_Array[85] := -126.566864, FeedBagVolume_Array[86] := -126.566864, FeedBagVolume_Array[87] := -126.566864, FeedBagVolume_Array[88] := -126.566864, FeedBagVolume_Array[89] := -126.566864, FeedBagVolume_Array[90] := -126.566864, FeedBagVolume_Array[91] := -126.566864, FeedBagVolume_Array[92] := -126.566864, FeedBagVolume_Array[93] := -126.566864, FeedBagVolume_Array[94] := -126.566864, FeedBagVolume_Array[95] := -126.566864, FeedBagVolume_Array[96] := -126.566864, FeedBagVolume_Array[97] := -126.566864, FeedBagVolume_Array[98] := -126.566864, FeedBagVolume_Array[99] := -126.566864, FeedBagVolume_Array[100] := -126.566864, FeedBagVolume_MAVE.In := -126.566864, FeedBagVolume_MAVE.SampleEnable := 1, FeedBagVolume_MAVE.NumberOfSamples := 1, FeedBagVolume_MAVE.Out := -126.566864, WI201_Unfiltered := -499.96185, FiltrateVolume := -495.01175, FiltrateVolume_Array[0] := -494.9362, FiltrateVolume_Array[1] := -495.01175, FiltrateVolume_Array[2] := -495.01175, FiltrateVolume_Array[3] := -495.01175, FiltrateVolume_Array[4] := -495.01175,
        FiltrateVolume_Array[5] := -495.01175, FiltrateVolume_Array[6] := -495.01175, FiltrateVolume_Array[7] := -495.01175, FiltrateVolume_Array[8] := -495.01175, FiltrateVolume_Array[9] := -495.01175, FiltrateVolume_Array[10] := -495.01175, FiltrateVolume_Array[11] := -495.01175, FiltrateVolume_Array[12] := -495.01175, FiltrateVolume_Array[13] := -495.01175, FiltrateVolume_Array[14] := -495.01175, FiltrateVolume_Array[15] := -495.01175, FiltrateVolume_Array[16] := -495.01175, FiltrateVolume_Array[17] := -495.01175, FiltrateVolume_Array[18] := -495.01175, FiltrateVolume_Array[19] := -495.01175, FiltrateVolume_Array[20] := -495.01175, FiltrateVolume_Array[21] := -494.9362, FiltrateVolume_Array[22] := -495.01175, FiltrateVolume_Array[23] := -495.01175, FiltrateVolume_Array[24] := -495.01175, FiltrateVolume_Array[25] := -495.01175, FiltrateVolume_Array[26] := -495.01175, FiltrateVolume_Array[27] := -495.01175, FiltrateVolume_Array[28] := -495.01175, FiltrateVolume_Array[29] := -495.01175, FiltrateVolume_Array[30] := -495.01175, FiltrateVolume_Array[31] := -495.01175, FiltrateVolume_Array[32] := -495.01175, FiltrateVolume_Array[33] := -495.01175, FiltrateVolume_Array[34] := -494.9362, FiltrateVolume_Array[35] := -494.9362, FiltrateVolume_Array[36] := -495.01175, FiltrateVolume_Array[37] := -495.01175, FiltrateVolume_Array[38] := -495.01175, FiltrateVolume_Array[39] := -495.01175, FiltrateVolume_Array[40] := -495.01175, FiltrateVolume_Array[41] := -495.01175, FiltrateVolume_Array[42] := -495.01175, FiltrateVolume_Array[43] := -494.9362, FiltrateVolume_Array[44] := -495.01175, FiltrateVolume_Array[45] := -494.9362, FiltrateVolume_Array[46] := -495.01175, FiltrateVolume_Array[47] := -495.01175, FiltrateVolume_Array[48] := -495.01175, FiltrateVolume_Array[49] := -495.01175, FiltrateVolume_Array[50] := -495.01175, FiltrateVolume_Array[51] := -495.01175, FiltrateVolume_Array[52] := -495.01175, FiltrateVolume_Array[53] := -495.01175, FiltrateVolume_Array[54] := -495.01175, FiltrateVolume_Array[55] := -495.01175, FiltrateVolume_Array[56] := -495.01175, FiltrateVolume_Array[57] := -495.01175, FiltrateVolume_Array[58] := -495.01175, FiltrateVolume_Array[59] := -495.01175, FiltrateVolume_Array[60] := -495.01175, FiltrateVolume_Array[61] := -495.01175, FiltrateVolume_Array[62] := -494.9362, FiltrateVolume_Array[63] := -494.9362, FiltrateVolume_Array[64] := -495.01175,
        FiltrateVolume_Array[65] := -494.9362, FiltrateVolume_Array[66] := -495.01175, FiltrateVolume_Array[67] := -495.01175, FiltrateVolume_Array[68] := -495.01175, FiltrateVolume_Array[69] := -494.9362, FiltrateVolume_Array[70] := -494.9362, FiltrateVolume_Array[71] := -495.01175, FiltrateVolume_Array[72] := -495.01175, FiltrateVolume_Array[73] := -495.01175, FiltrateVolume_Array[74] := -495.01175, FiltrateVolume_Array[75] := -494.9362, FiltrateVolume_Array[76] := -495.01175, FiltrateVolume_Array[77] := -495.01175, FiltrateVolume_Array[78] := -495.01175, FiltrateVolume_Array[79] := -495.01175, FiltrateVolume_Array[80] := -495.01175, FiltrateVolume_Array[81] := -495.01175, FiltrateVolume_Array[82] := -495.01175, FiltrateVolume_Array[83] := -495.01175, FiltrateVolume_Array[84] := -495.01175, FiltrateVolume_Array[85] := -495.01175, FiltrateVolume_Array[86] := -495.01175, FiltrateVolume_Array[87] := -495.01175, FiltrateVolume_Array[88] := -495.01175, FiltrateVolume_Array[89] := -495.01175, FiltrateVolume_Array[90] := -495.01175, FiltrateVolume_Array[91] := -495.01175, FiltrateVolume_Array[92] := -495.01175, FiltrateVolume_Array[93] := -495.01175, FiltrateVolume_Array[94] := -495.01175, FiltrateVolume_Array[95] := -495.01175, FiltrateVolume_Array[96] := -494.9362, FiltrateVolume_Array[97] := -495.01175, FiltrateVolume_Array[98] := -495.01175, FiltrateVolume_Array[99] := -495.01175, FiltrateVolume_Array[100] := -495.01175, FiltrateVolume_MAVE.In := -495.01175, FiltrateVolume_MAVE.SampleEnable := 1, FiltrateVolume_MAVE.NumberOfSamples := 1, FiltrateVolume_MAVE.Out := -495.01175, FiltrateVolume_MaveFiltered := -495.01175, FiltrateVolume_ExpConst := 0.99, FiltrateVolume_ExpFiltered := -495.0009, Weight_ExpFiltered := -499.9509, Weight_MaveFiltered := -499.96185);   // Data for Scale Filtering
   SIC001 : ALIAS FOR Drive[1];
   SIC001_AO : ALIAS FOR AnalogOutput[0];
   SIC001_DO : ALIAS FOR DigitalOutput[8];
   SIC001DF : ALIAS FOR DigitalPoint[16];
   SIC002 : ALIAS FOR Drive[2];
   SIC002_AO : ALIAS FOR AnalogOutput[1];
   SIC002_DO : ALIAS FOR DigitalOutput[9];
   SIC002DF : ALIAS FOR DigitalPoint[17];
   SIC003_AO : ALIAS FOR AnalogOutput[2];
   SIC003_DO : ALIAS FOR DigitalOutput[15];
   SIC003DF : ALIAS FOR DigitalPoint[29];
   SIC004 : ALIAS FOR Drive[3];
   SIC004_AO : ALIAS FOR AnalogOutput[5];
   SysControl : SysControl := (DefaultTimer.PRE := 3000, AllAutoTimer.PRE := 3000, DefaultStatus := 1, EnableSaveRestoreParam := 1, UV_Auto_Zero_Timer.PRE := 3000, Tare_WI101_Timer.PRE := 3000, ClearTare_WI101_Timer.PRE := 3000, Zero_WI101_Timer.PRE := 3000, Tare_PI001_Timer.PRE := 3000, Tare_PI101_Timer.PRE := 3000, Tare_PI201_Timer.PRE := 3000, Tare_PI401_Timer.PRE := 3000, Tare_PI601_Timer.PRE := 3000);   // General system status and command
   Tank : TankManagement := (Config.TankSelected := 4, Config.TankSelectHMI := 500, Config.TankSelectPLC := 500, Config.Option_Prev := 4, Config.TMR.PRE := 500, WeightConfiguration[0].Alm_HI := 2.0, WeightConfiguration[0].Alm_HI_PRE := 2.0, WeightConfiguration[0].Alm_HIHI := 2.0, WeightConfiguration[0].Alm_HIHI_PRE := 2.0, WeightConfiguration[0].Alm_LOLOTMR := 2, WeightConfiguration[0].Alm_LOLOTMR_PRE := 2, WeightConfiguration[0].Alm_LOTMR := 2, WeightConfiguration[0].Alm_LOTMR_PRE := 2, WeightConfiguration[0].Alm_HITMR := 2, WeightConfiguration[0].Alm_HITMR_PRE := 2, WeightConfiguration[0].Alm_HIHITMR := 2, WeightConfiguration[0].Alm_HIHITMR_PRE := 2, WeightConfiguration[1].Desc := '50L', WeightConfiguration[1].Alm_HI := 50.0, WeightConfiguration[1].Alm_HI_PRE := 50.0, WeightConfiguration[1].Alm_HIHI := 50.0, WeightConfiguration[1].Alm_HIHI_PRE := 50.0, WeightConfiguration[1].Alm_LOLOTMR := 5, WeightConfiguration[1].Alm_LOLOTMR_PRE := 5, WeightConfiguration[1].Alm_LOTMR := 2, WeightConfiguration[1].Alm_LOTMR_PRE := 2, WeightConfiguration[1].Alm_HITMR := 2, WeightConfiguration[1].Alm_HITMR_PRE := 2, WeightConfiguration[1].Alm_HIHITMR := 5, WeightConfiguration[1].Alm_HIHITMR_PRE := 5, WeightConfiguration[2].Desc := '100L', WeightConfiguration[2].Alm_HI := 100.0, WeightConfiguration[2].Alm_HI_PRE := 100.0, WeightConfiguration[2].Alm_HIHI := 100.0, WeightConfiguration[2].Alm_HIHI_PRE := 100.0, WeightConfiguration[2].Alm_LOLOTMR := 5, WeightConfiguration[2].Alm_LOLOTMR_PRE := 5, WeightConfiguration[2].Alm_LOTMR := 2, WeightConfiguration[2].Alm_LOTMR_PRE := 2, WeightConfiguration[2].Alm_HITMR := 2, WeightConfiguration[2].Alm_HITMR_PRE := 2, WeightConfiguration[2].Alm_HIHITMR := 5, WeightConfiguration[2].Alm_HIHITMR_PRE := 5, WeightConfiguration[3].Desc := '200L', WeightConfiguration[3].Alm_HI := 240.0, WeightConfiguration[3].Alm_HI_PRE := 240.0, WeightConfiguration[3].Alm_HIHI := 240.0, WeightConfiguration[3].Alm_HIHI_PRE := 240.0, WeightConfiguration[3].Alm_LOLOTMR := 2, WeightConfiguration[3].Alm_LOLOTMR_PRE := 2, WeightConfiguration[3].Alm_LOTMR := 2, WeightConfiguration[3].Alm_LOTMR_PRE := 2, WeightConfiguration[3].Alm_HITMR := 2, WeightConfiguration[3].Alm_HITMR_PRE := 2, WeightConfiguration[3].Alm_HIHITMR := 2, WeightConfiguration[3].Alm_HIHITMR_PRE := 2, WeightConfiguration[4].Desc := '500L', WeightConfiguration[4].Alm_LOLO := 105.0, WeightConfiguration[4].Alm_LOLO_PRE := 105.0, WeightConfiguration[4].Alm_LO := 110.0,
        WeightConfiguration[4].Alm_LO_PRE := 110.0, WeightConfiguration[4].Alm_HI := 400.0, WeightConfiguration[4].Alm_HI_PRE := 400.0, WeightConfiguration[4].Alm_HIHI := 450.0, WeightConfiguration[4].Alm_HIHI_PRE := 450.0, WeightConfiguration[4].Alm_LOLOTMR := 2, WeightConfiguration[4].Alm_LOLOTMR_PRE := 2, WeightConfiguration[4].Alm_LOTMR := 2, WeightConfiguration[4].Alm_LOTMR_PRE := 2, WeightConfiguration[4].Alm_HITMR := 2, WeightConfiguration[4].Alm_HITMR_PRE := 2, WeightConfiguration[4].Alm_HIHITMR := 2, WeightConfiguration[4].Alm_HIHITMR_PRE := 2, LevelConfiguration[0].Alm_HI := 99999.0, LevelConfiguration[0].Alm_HI_PRE := 99999.0, LevelConfiguration[0].Alm_HIHI := 99999.0, LevelConfiguration[0].Alm_HIHI_PRE := 99999.0, LevelConfiguration[0].Alm_LOLOTMR := 2, LevelConfiguration[0].Alm_LOLOTMR_PRE := 2, LevelConfiguration[0].Alm_LOTMR := 2, LevelConfiguration[0].Alm_LOTMR_PRE := 2, LevelConfiguration[0].Alm_HITMR := 2, LevelConfiguration[0].Alm_HITMR_PRE := 2, LevelConfiguration[0].Alm_HIHITMR := 2, LevelConfiguration[0].Alm_HIHITMR_PRE := 2, LevelConfiguration[1].Desc := '50L', LevelConfiguration[1].ScaledMax := 50.0, LevelConfiguration[1].ScaledMax_PRE := 50.0, LevelConfiguration[1].Alm_HI := 50.0, LevelConfiguration[1].Alm_HI_PRE := 50.0, LevelConfiguration[1].Alm_HIHI := 50.0, LevelConfiguration[1].Alm_HIHI_PRE := 50.0, LevelConfiguration[1].Alm_LOLOTMR := 5, LevelConfiguration[1].Alm_LOLOTMR_PRE := 5, LevelConfiguration[1].Alm_LOTMR := 2, LevelConfiguration[1].Alm_LOTMR_PRE := 2, LevelConfiguration[1].Alm_HITMR := 2, LevelConfiguration[1].Alm_HITMR_PRE := 2, LevelConfiguration[1].Alm_HIHITMR := 5, LevelConfiguration[1].Alm_HIHITMR_PRE := 5, LevelConfiguration[2].Desc := '100L', LevelConfiguration[2].ScaledMax := 100.0, LevelConfiguration[2].ScaledMax_PRE := 100.0, LevelConfiguration[2].Alm_HI := 100.0, LevelConfiguration[2].Alm_HI_PRE := 100.0, LevelConfiguration[2].Alm_HIHI := 100.0, LevelConfiguration[2].Alm_HIHI_PRE := 100.0, LevelConfiguration[2].Alm_LOLOTMR := 5, LevelConfiguration[2].Alm_LOLOTMR_PRE := 5, LevelConfiguration[2].Alm_LOTMR := 2, LevelConfiguration[2].Alm_LOTMR_PRE := 2, LevelConfiguration[2].Alm_HITMR := 2, LevelConfiguration[2].Alm_HITMR_PRE := 2, LevelConfiguration[2].Alm_HIHITMR := 5, LevelConfiguration[2].Alm_HIHITMR_PRE := 5, LevelConfiguration[3].Desc := '200L', LevelConfiguration[3].ScaledMax := 200.0, LevelConfiguration[3].ScaledMax_PRE := 200.0, LevelConfiguration[3].Alm_HI := 200.0, LevelConfiguration[3].Alm_HI_PRE := 200.0,
        LevelConfiguration[3].Alm_HIHI := 200.0, LevelConfiguration[3].Alm_HIHI_PRE := 200.0, LevelConfiguration[3].Alm_LOLOTMR := 2, LevelConfiguration[3].Alm_LOLOTMR_PRE := 2, LevelConfiguration[3].Alm_LOTMR := 2, LevelConfiguration[3].Alm_LOTMR_PRE := 2, LevelConfiguration[3].Alm_HITMR := 2, LevelConfiguration[3].Alm_HITMR_PRE := 2, LevelConfiguration[3].Alm_HIHITMR := 2, LevelConfiguration[3].Alm_HIHITMR_PRE := 2, LevelConfiguration[4].Desc := '500L', LevelConfiguration[4].ScaledMax := 500.0, LevelConfiguration[4].ScaledMax_PRE := 500.0, LevelConfiguration[4].Alm_LOLO := 90.0, LevelConfiguration[4].Alm_LOLO_PRE := 90.0, LevelConfiguration[4].Alm_LO := 100.0, LevelConfiguration[4].Alm_LO_PRE := 100.0, LevelConfiguration[4].Alm_HI := 200.0, LevelConfiguration[4].Alm_HI_PRE := 200.0, LevelConfiguration[4].Alm_HIHI := 300.0, LevelConfiguration[4].Alm_HIHI_PRE := 300.0, LevelConfiguration[4].Alm_LOLOTMR := 2, LevelConfiguration[4].Alm_LOLOTMR_PRE := 2, LevelConfiguration[4].Alm_LOTMR := 2, LevelConfiguration[4].Alm_LOTMR_PRE := 2, LevelConfiguration[4].Alm_HITMR := 2, LevelConfiguration[4].Alm_HITMR_PRE := 2, LevelConfiguration[4].Alm_HIHITMR := 2, LevelConfiguration[4].Alm_HIHITMR_PRE := 2);   // Tank Management
   TCU101 : ALIAS FOR AnalogPoint[18];
   TCU101_AO : ALIAS FOR AnalogOutput[6];
   TCU101_SIG : ALIAS FOR DigitalPoint[108];
   TCU101Alarm : ALIAS FOR AlarmAnalog[18];
   TCU101DF : ALIAS FOR DigitalPoint[30];
   TCU101ON : ALIAS FOR DigitalOutput[20];
   ThisSystem : SystemType := (Value := 2, MoldType := 126, PreviousValue := 126, EnableSystemType[0] := 1, EnableSystemType[3] := 1, NewSystem_Timer.PRE := 60000, NewSystem_Timer.ACC := 177455, NewSystem_Timer.EN := 1, NewSystem_Timer.DN := 1);
   TI101 : ALIAS FOR AnalogPoint[13];
   TI101_SIG : ALIAS FOR DigitalPoint[101];
   TI101Alarm : ALIAS FOR AlarmAnalog[13];
   TI201 : ALIAS FOR AnalogPoint[22];
   TI201_SIG : ALIAS FOR DigitalPoint[111];
   TI201Alarm : ALIAS FOR AlarmAnalog[22];
   TIC101Control : TCUControl := (SP_Disable := 20.0, Offset := 15.0, OffsetTimer.PRE := 30000, OffsetTime := 30.0, LevelMin := 20.0);
   TimerControl : TimerControl := (TickMainTask := 1, Save := 18526, Seconds := 18526, Colon := ':', ColonZero := ':0', Cycle := 741044);   // Timer Control
   Timers : Timers[22] := ([0].TotalSeconds := 44.0, [0].Seconds := 44, [0].sHours := '0', [0].sMinutes := '0', [0].sSeconds := '44', [0].HMS := '0:00:44', [0].LastHMS := '0:02:09', [1].TotalSeconds := 21.0, [1].Seconds := 21, [1].sHours := '0', [1].sMinutes := '0', [1].sSeconds := '21', [1].HMS := '0:00:21', [2].TotalSeconds := 1.0, [2].Seconds := 1, [2].sHours := '0', [2].sMinutes := '0', [2].sSeconds := '1', [2].HMS := '0:00:01', [3].TotalSeconds := 9.0, [3].Seconds := 9, [3].sHours := '0', [3].sMinutes := '0', [3].sSeconds := '9', [3].HMS := '0:00:09', [3].LastHMS := '0:00:00', [4].sHours := '0', [4].sMinutes := '0', [4].sSeconds := '0', [4].HMS := '0:00:00', [5].sHours := '0', [5].sMinutes := '0', [5].sSeconds := '0', [5].HMS := '0:00:00', [5].LastHMS := ':00$00$07$00$00$000:00:00$00$00$00$00$00$00$00$00$00$07$00$00$00', [6].TotalSeconds := 9.0, [6].Seconds := 9, [6].sHours := '0', [6].sMinutes := '0', [6].sSeconds := '9', [6].HMS := '0:00:09', [6].LastHMS := '0:00:02', [7].sHours := '0', [7].sMinutes := '0', [7].sSeconds := '0', [7].HMS := '0:00:00', [8].sHours := '0', [8].sMinutes := '0', [8].sSeconds := '0', [8].HMS := '0:00:00', [8].LastHMS := '$07$00$00$000:00:00$00$00$00$00$00$00$00$00$00$07$00$00$000:$00$00', [9].TotalSeconds := 2.0, [9].Seconds := 2, [9].sHours := '0', [9].sMinutes := '0', [9].sSeconds := '2', [9].HMS := '0:00:02', [9].LastHMS := '$00$00$00$00$00$00$00$00$07$00$00$000:00:00$00$07$00$00$000:$00$00', [10].sHours := '0', [10].sMinutes := '0',
        [10].sSeconds := '0', [10].HMS := '0:00:00', [10].LastHMS := '0:00:00', [11].sHours := '0', [11].sMinutes := '0', [11].sSeconds := '0', [11].HMS := '0:00:00', [11].LastHMS := '0:00:00', [12].sHours := '0', [12].sMinutes := '0', [12].sSeconds := '0', [12].HMS := '0:00:00', [13].sHours := '0', [13].sMinutes := '0', [13].sSeconds := '0', [13].HMS := '0:00:00', [13].LastHMS := ':00$00$07$00$00$000:00:00$00$00$00$00$00$00$00$00$00$07$00$00$00', [14].sHours := '0', [14].sMinutes := '0', [14].sSeconds := '0', [14].HMS := '0:00:00', [14].LastHMS := ':00$00$00$00$00$00$00$00$00$00$07$00$00$000:00:00$00$07$00$00$00', [15].sHours := '0', [15].sMinutes := '0', [15].sSeconds := '0', [15].HMS := '0:00:00', [16].sHours := '0', [16].sMinutes := '0', [16].sSeconds := '0', [16].HMS := '0:00:00', [16].LastHMS := '$07$00$00$000:00:00$00$00$00$00$00$00$00$00$00$07$00$00$000:$00$00', [17].sHours := '0', [17].sMinutes := '0', [17].sSeconds := '0', [17].HMS := '0:00:00', [17].LastHMS := '$00$00$00$00$00$00$00$00$07$00$00$000:00:00$00$07$00$00$000:$00$00', [18].sHours := '0', [18].sMinutes := '0', [18].sSeconds := '0', [18].HMS := '0:00:00', [18].LastHMS := '0:00:00', [19].TotalSeconds := 49.0, [19].Seconds := 49, [19].sHours := '0', [19].sMinutes := '0', [19].sSeconds := '49', [19].HMS := '0:00:49', [19].LastHMS := '0:00:00', [20].Enable := 1, [20].TotalSeconds := 427.0, [20].Minutes := 7, [20].Seconds := 7, [20].sHours := '0', [20].sMinutes := '7', [20].sSeconds := '7', [20].HMS := '0:07:07', [21].sHours := '0', [21].sMinutes := '0', [21].sSeconds := '0', [21].HMS := '0:00:00',
        [21].LastHMS := '0:00:00');   // Timer Array
        [10]   // Phase 4 Step Time
        [19]   // Procedure Time
        [0]   // Phase 0 Total Time
        [11]   // Phase 5 Step Time
        [12]   // Phase 0 Pause Time
        [13]   // Phase 1 Pause Time
        [14]   // Phase 2 Pause Time
        [15]   // Phase 3 Pause Time
        [16]   // Phase 4 Pause Time
        [17]   // Phase 5 Pause Time
        [18]   // User Time
        [1]   // Phase 1 Total Time
        [21]   // Linear Gradient
        [2]   // Phase 2 Total Time
        [3]   // Phase 3 Total Time
        [4]   // Phase 4 Total Time
        [5]   // Phase 5 Total Time
        [6]   // Phase 0 Step Time
        [7]   // Phase 1 Step Time
        [8]   // Phase 2 Step Time
        [9]   // Phase 3 Step Time
   TMP : ALIAS FOR AnalogPoint[41];
   TMPAlarm : ALIAS FOR AlarmAnalog[41];
   TNK101 : ALIAS FOR DigitalOutput[18];
   TNK102 : ALIAS FOR DigitalOutput[19];
   TNK103 : ALIAS FOR DigitalOutput[27];
   Totalizer : Totalizers[20] := ([0].PV := -23.769741, [0].PVscale := 60.0, [0].Title := 'Conc', [0].ResetTimer.PRE := 3000, [1].PV := -23.769741, [1].PVscale := 60.0, [1].Title := 'Diaf', [1].ResetTimer.PRE := 3000, [2].ResetTimer.PRE := 3000, [3].ResetTimer.PRE := 3000, [4].ResetTimer.PRE := 3000, [5].ResetTimer.PRE := 3000, [6].ResetTimer.PRE := 3000, [7].ResetTimer.PRE := 3000, [8].ResetTimer.PRE := 3000, [9].ResetTimer.PRE := 3000, [10].ResetTimer.PRE := 3000, [11].ResetTimer.PRE := 3000, [12].ResetTimer.PRE := 3000, [13].ResetTimer.PRE := 3000, [14].ResetTimer.PRE := 3000, [15].ResetTimer.PRE := 3000, [16].ResetTimer.PRE := 3000, [17].ResetTimer.PRE := 3000, [18].ResetTimer.PRE := 3000, [19].ResetTimer.PRE := 3000);   // Totalizers Array
        [0]   // Concentration totalizer
        [1]   // Diafiltration totalizer
   UserAlarm : UserAlarm;   // User Alarm (used in CCP Recipe)
   UserCr1 : ALIAS FOR DigitalPoint[65];
   UserCr2 : ALIAS FOR DigitalPoint[67];
   UserNCr1 : ALIAS FOR DigitalPoint[64];
   UserNCr2 : ALIAS FOR DigitalPoint[66];
   UserTime : ALIAS FOR Timers[18];   // User time
   UserTotalizerManagement : UserTotalizerManagement := (LogUserTimer.PRE := 3000, ResetUserTimer.PRE := 3000);   // User Totalizer management
   Valve : Valve[100] := ([0].Tag := 'XV001', [0].Control := 1, [0].Auto := 1, [0].Manual := 1, [0].OpenStatus := 1, [0].ZSOverride := 1, [0].FailState := 1, [0].EnableCfg := 1, [0].StatusWord := 2, [0].Status := 2, [0].OutputAddress := 32, [0].AlarmTimer.PRE := 2000, [0].AlarmTimerSP := 2, [1].Tag := 'XV002', [1].Control := 1, [1].Auto := 1, [1].Manual := 1, [1].OpenStatus := 1, [1].ZSOverride := 1, [1].FailState := 1, [1].EnableCfg := 1, [1].StatusWord := 2, [1].Status := 2, [1].OutputAddress := 33, [1].AlarmTimer.PRE := 2000, [1].AlarmTimerSP := 2, [1].AutoCloseTimer.ACC := 1103, [2].Tag := 'XV003', [2].ZSOpenEnable := 1, [2].CloseStatus := 1, [2].ZSOverride := 1, [2].PriorityCfg := 1, [2].EnableCfg := 1, [2].StatusWord := 4, [2].Status := 4, [2].ZSOpenAddress := 2, [2].OutputAddress := 34, [2].AlarmTimer.PRE := 2000, [2].AlarmTimerSP := 2, [2].AutoCloseTimer.ACC := 1032, [3].Tag := 'XV004', [3].ZSOpenEnable := 1, [3].CloseStatus := 1, [3].ZSOverride := 1, [3].PriorityCfg := 1, [3].EnableCfg := 1, [3].StatusWord := 4, [3].Status := 4, [3].ZSOpenAddress := 3, [3].OutputAddress := 35, [3].AlarmTimer.PRE := 2000, [3].AlarmTimerSP := 2, [3].AutoCloseTimer.ACC := 1115, [4].Tag := 'XV005', [4].ZSOpenEnable := 1, [4].CloseStatus := 1, [4].ZSOverride := 1, [4].PriorityCfg := 1, [4].EnableCfg := 1, [4].StatusWord := 4,
        [4].Status := 4, [4].ZSOpenAddress := 4, [4].OutputAddress := 36, [4].AlarmTimer.PRE := 2000, [4].AlarmTimerSP := 2, [4].AutoCloseTimer.ACC := 1104, [5].Tag := 'XV102', [5].ZSOpenEnable := 1, [5].CloseStatus := 1, [5].ZSOverride := 1, [5].PriorityCfg := 1, [5].EnableCfg := 1, [5].StatusWord := 4, [5].Status := 4, [5].ZSOpenAddress := 5, [5].OutputAddress := 37, [5].AlarmTimer.PRE := 2000, [5].AlarmTimerSP := 2, [5].AutoCloseTimer.ACC := 1104, [6].Tag := 'XV401', [6].ZSOpenEnable := 1, [6].CloseStatus := 1, [6].ZSOverride := 1, [6].PriorityCfg := 1, [6].EnableCfg := 1, [6].StatusWord := 4, [6].Status := 4, [6].ZSOpenAddress := 6, [6].OutputAddress := 38, [6].AlarmTimer.PRE := 2000, [6].AlarmTimerSP := 2, [6].AutoCloseTimer.ACC := 1104, [7].Tag := 'XV402', [7].Control := 1, [7].Auto := 1, [7].Manual := 1, [7].OpenStatus := 1, [7].ZSOverride := 1, [7].FailState := 1, [7].EnableCfg := 1, [7].StatusWord := 2, [7].Status := 2, [7].OutputAddress := 39, [7].AlarmTimer.PRE := 2000, [7].AlarmTimerSP := 2, [7].AutoCloseTimer.ACC := 1104, [8].Tag := 'XV411', [8].Control := 1, [8].Auto := 1, [8].Manual := 1, [8].OpenStatus := 1, [8].ZSOverride := 1, [8].FailState := 1, [8].EnableCfg := 1, [8].StatusWord := 2, [8].Status := 2, [8].OutputAddress := 40, [8].AlarmTimer.PRE := 2000, [8].AlarmTimerSP := 2, [8].AutoCloseTimer.ACC := 1104,
        [9].Tag := 'XV421', [9].CloseStatus := 1, [9].ZSOverride := 1, [9].EnableCfg := 1, [9].StatusWord := 4, [9].Status := 4, [9].OutputAddress := 41, [9].AlarmTimer.PRE := 2000, [9].AlarmTimerSP := 2, [9].AutoCloseTimer.ACC := 1105, [10].Tag := 'XV431', [10].CloseStatus := 1, [10].ZSOverride := 1, [10].EnableCfg := 1, [10].StatusWord := 4, [10].Status := 4, [10].OutputAddress := 42, [10].AlarmTimer.PRE := 2000, [10].AlarmTimerSP := 2, [10].AutoCloseTimer.ACC := 1104, [11].Tag := 'XV441', [11].CloseStatus := 1, [11].ZSOverride := 1, [11].EnableCfg := 1, [11].StatusWord := 4, [11].Status := 4, [11].OutputAddress := 43, [11].AlarmTimer.PRE := 2000, [11].AlarmTimerSP := 2, [11].AutoCloseTimer.ACC := 1103, [12].Tag := 'XV501', [12].CloseStatus := 1, [12].ZSOverride := 1, [12].EnableCfg := 1, [12].StatusWord := 4, [12].Status := 4, [12].OutputAddress := 44, [12].AlarmTimer.PRE := 2000, [12].AlarmTimerSP := 2, [12].AutoCloseTimer.ACC := 1072, [13].Tag := 'XV502', [13].CloseStatus := 1, [13].ZSOverride := 1, [13].StatusWord := 4, [13].Status := 4, [13].OutputAddress := 45, [13].AlarmTimer.PRE := 2000, [13].AlarmTimerSP := 2, [13].AutoCloseTimer.ACC := 1016, [14].Tag := 'XV901', [14].CloseStatus := 1, [14].ZSOverride := 1, [14].StatusWord := 4, [14].Status := 4, [14].OutputAddress := 46, [14].AlarmTimer.PRE := 2000, [14].AlarmTimerSP := 2, [15].CloseStatus := 1, [15].ZSOverride := 1, [15].EnableCfg := 1,
        [15].StatusWord := 4, [15].Status := 4, [15].OutputAddress := 47, [15].AlarmTimer.PRE := 2000, [15].AlarmTimerSP := 2, [16].CloseStatus := 1, [16].ZSOverride := 1, [16].EnableCfg := 1, [16].StatusWord := 4, [16].Status := 4, [16].OutputAddress := 48, [16].AlarmTimer.PRE := 2000, [16].AlarmTimerSP := 2, [17].CloseStatus := 1, [17].ZSOverride := 1, [17].EnableCfg := 1, [17].StatusWord := 4, [17].Status := 4, [17].OutputAddress := 49, [17].AlarmTimer.PRE := 2000, [17].AlarmTimerSP := 2, [17].AutoCloseTimer.ACC := 1594, [18].CloseStatus := 1, [18].ZSOverride := 1, [18].EnableCfg := 1, [18].StatusWord := 4, [18].Status := 4, [18].OutputAddress := 50, [18].AlarmTimer.PRE := 2000, [18].AlarmTimerSP := 2, [18].AutoCloseTimer.ACC := 137, [19].CloseStatus := 1, [19].ZSOverride := 1, [19].EnableCfg := 1, [19].StatusWord := 4, [19].Status := 4, [19].OutputAddress := 51, [19].AlarmTimer.PRE := 2000, [19].AlarmTimerSP := 2, [19].AutoCloseTimer.ACC := 1007, [20].CloseStatus := 1, [20].ZSOverride := 1, [20].EnableCfg := 1, [20].StatusWord := 4, [20].Status := 4, [20].OutputAddress := 52, [20].AlarmTimer.PRE := 2000, [20].AlarmTimerSP := 2, [20].AutoCloseTimer.ACC := 1004, [21].OpenStatus := 1, [21].AlarmTimerSP := 2, [22].CloseStatus := 1, [22].AlarmTimerSP := 2, [22].AutoCloseTimer.ACC := 131, [23].CloseStatus := 1, [23].AlarmTimerSP := 2, [23].AutoCloseTimer.ACC := 1003, [24].CloseStatus := 1, [24].AlarmTimerSP := 2, [24].AutoCloseTimer.ACC := 1002,
        [25].CloseStatus := 1, [25].AlarmTimerSP := 2, [25].AutoCloseTimer.ACC := 1002, [26].CloseStatus := 1, [26].AlarmTimerSP := 2, [26].AutoCloseTimer.ACC := 1002, [27].CloseStatus := 1, [27].AlarmTimerSP := 2, [28].CloseStatus := 1, [28].AlarmTimerSP := 2, [29].OpenStatus := 1, [29].AlarmTimerSP := 2, [29].AutoCloseTimer.ACC := 1068, [30].CloseStatus := 1, [30].AlarmTimerSP := 2, [30].AutoCloseTimer.ACC := 1069, [31].CloseStatus := 1, [31].AlarmTimerSP := 2, [31].AutoCloseTimer.ACC := 131, [32].CloseStatus := 1, [32].PriorityCfg := 1, [32].AlarmTimerSP := 2, [32].AutoCloseTimer.ACC := 1059, [33].OpenStatus := 1, [33].PriorityCfg := 1, [33].AlarmTimerSP := 2, [33].AutoCloseTimer.ACC := 1123, [34].OpenStatus := 1, [34].PriorityCfg := 1, [34].AlarmTimerSP := 2, [34].AutoCloseTimer.ACC := 1095, [35].OpenStatus := 1, [35].PriorityCfg := 1, [35].AlarmTimerSP := 2, [35].AutoCloseTimer.ACC := 1127, [36].OpenStatus := 1, [36].PriorityCfg := 1, [36].AlarmTimerSP := 2, [36].AutoCloseTimer.ACC := 1004, [37].CloseStatus := 1, [37].PriorityCfg := 1, [37].AlarmTimerSP := 2, [37].AutoCloseTimer.ACC := 1121, [38].CloseStatus := 1, [38].Priority := 1, [38].PriorityCfg := 1, [38].AlarmTimerSP := 2, [38].AutoCloseTimer.ACC := 1135, [39].CloseStatus := 1, [39].Priority := 1, [39].PriorityCfg := 1, [39].AlarmTimerSP := 2, [39].AutoCloseTimer.ACC := 1121, [40].CloseStatus := 1, [40].Priority := 1, [40].PriorityCfg := 1, [40].AlarmTimerSP := 2, [40].AutoCloseTimer.ACC := 1112, [41].CloseStatus := 1, [41].Priority := 1,
        [41].PriorityCfg := 1, [41].AlarmTimerSP := 2, [42].CloseStatus := 1, [42].Priority := 1, [42].PriorityCfg := 1, [42].AlarmTimerSP := 2, [43].CloseStatus := 1, [43].Priority := 1, [43].PriorityCfg := 1, [43].AlarmTimerSP := 2, [44].CloseStatus := 1, [44].Priority := 1, [44].PriorityCfg := 1, [44].AlarmTimerSP := 2, [45].CloseStatus := 1, [45].Priority := 1, [45].PriorityCfg := 1, [45].AlarmTimerSP := 2, [46].CloseStatus := 1, [46].Priority := 1, [46].PriorityCfg := 1, [46].AlarmTimerSP := 2, [47].OpenStatus := 1, [47].Priority := 1, [47].PriorityCfg := 1, [47].AlarmTimerSP := 2, [51].OpenStatus := 1, [52].OpenStatus := 1, [53].CloseStatus := 1, [54].CloseStatus := 1, [55].CloseStatus := 1, [56].CloseStatus := 1, [58].CloseStatus := 1, [59].CloseStatus := 1);   // Valve Array
        [10]   // XV402
        [11]   // XV403
        [12]   // XV404
        [0]   // XV001
        [0].FailState   // Valve Fail State 0=Closed 1=Open
        [13]   // XV405
        [14]   // XV406
        [15]   // XV201
        [16]   // XV202
        [17]   // XV701
        [18]   // XV702
        [19]   // XV703
        [20]   // XV704
        [1]   // XV002
        [2]   // XV003
        [3]   // XV004
        [4]   // XV005
        [5]   // XV006
        [6]   // XV007
        [7]   // XV101
        [8]   // XV102
        [9]   // XV401
   Valve_Storage : Valve[6,100] := ([0,0].Tag := 'XV001', [0,0].CloseStatus := 1, [0,0].ZSOverride := 1, [0,0].EnableCfg := 1, [0,0].StatusWord := 4, [0,0].Status := 4, [0,0].OutputAddress := 32, [0,0].AlarmTimer.PRE := 2000, [0,0].AlarmTimerSP := 2, [0,1].Tag := 'XV002', [0,1].CloseStatus := 1, [0,1].ZSOverride := 1, [0,1].EnableCfg := 1, [0,1].StatusWord := 4, [0,1].Status := 4, [0,1].OutputAddress := 33, [0,1].AlarmTimer.PRE := 2000, [0,1].AlarmTimerSP := 2, [0,1].AutoCloseTimer.ACC := 1103, [0,2].Tag := 'XV003', [0,2].CloseStatus := 1, [0,2].ZSOverride := 1, [0,2].EnableCfg := 1, [0,2].StatusWord := 4, [0,2].Status := 4, [0,2].OutputAddress := 34, [0,2].AlarmTimer.PRE := 2000, [0,2].AlarmTimerSP := 2, [0,2].AutoCloseTimer.ACC := 1032, [0,3].Tag := 'XV004', [0,3].CloseStatus := 1, [0,3].ZSOverride := 1, [0,3].EnableCfg := 1, [0,3].StatusWord := 4, [0,3].Status := 4, [0,3].OutputAddress := 35, [0,3].AlarmTimer.PRE := 2000, [0,3].AlarmTimerSP := 2, [0,3].AutoCloseTimer.ACC := 1115, [0,4].Tag := 'XV005', [0,4].CloseStatus := 1, [0,4].ZSOverride := 1, [0,4].EnableCfg := 1, [0,4].StatusWord := 4, [0,4].Status := 4, [0,4].OutputAddress := 36, [0,4].AlarmTimer.PRE := 2000, [0,4].AlarmTimerSP := 2, [0,4].AutoCloseTimer.ACC := 1104, [0,5].Tag := 'XV006', [0,5].CloseStatus := 1, [0,5].ZSOverride := 1, [0,5].EnableCfg := 1, [0,5].StatusWord := 4, [0,5].Status := 4, [0,5].OutputAddress := 37, [0,5].AlarmTimer.PRE := 2000, [0,5].AlarmTimerSP := 2, [0,5].AutoCloseTimer.ACC := 1104, [0,6].Tag := 'XV007',
        [0,6].CloseStatus := 1, [0,6].ZSOverride := 1, [0,6].EnableCfg := 1, [0,6].StatusWord := 4, [0,6].Status := 4, [0,6].OutputAddress := 38, [0,6].AlarmTimer.PRE := 2000, [0,6].AlarmTimerSP := 2, [0,6].AutoCloseTimer.ACC := 1104, [0,7].Tag := 'XV008', [0,7].CloseStatus := 1, [0,7].ZSOverride := 1, [0,7].EnableCfg := 1, [0,7].StatusWord := 4, [0,7].Status := 4, [0,7].OutputAddress := 39, [0,7].AlarmTimer.PRE := 2000, [0,7].AlarmTimerSP := 2, [0,7].AutoCloseTimer.ACC := 1104, [0,8].Tag := 'XV009', [0,8].CloseStatus := 1, [0,8].ZSOverride := 1, [0,8].EnableCfg := 1, [0,8].StatusWord := 4, [0,8].Status := 4, [0,8].OutputAddress := 40, [0,8].AlarmTimer.PRE := 2000, [0,8].AlarmTimerSP := 2, [0,8].AutoCloseTimer.ACC := 1104, [0,9].Tag := 'XV010', [0,9].CloseStatus := 1, [0,9].ZSOverride := 1, [0,9].EnableCfg := 1, [0,9].StatusWord := 4, [0,9].Status := 4, [0,9].OutputAddress := 41, [0,9].AlarmTimer.PRE := 2000, [0,9].AlarmTimerSP := 2, [0,9].AutoCloseTimer.ACC := 1105, [0,10].Tag := 'XV011', [0,10].CloseStatus := 1, [0,10].ZSOverride := 1, [0,10].EnableCfg := 1, [0,10].StatusWord := 4, [0,10].Status := 4, [0,10].OutputAddress := 42, [0,10].AlarmTimer.PRE := 2000, [0,10].AlarmTimerSP := 2, [0,10].AutoCloseTimer.ACC := 1104, [0,11].Tag := 'XV012', [0,11].Control := 1, [0,11].Auto := 1, [0,11].Manual := 1, [0,11].OpenStatus := 1, [0,11].ZSOverride := 1, [0,11].FailState := 1, [0,11].EnableCfg := 1, [0,11].StatusWord := 2, [0,11].Status := 2, [0,11].OutputAddress := 43,
        [0,11].AlarmTimer.PRE := 2000, [0,11].AlarmTimerSP := 2, [0,11].AutoCloseTimer.ACC := 1103, [0,12].Tag := 'XV013', [0,12].Control := 1, [0,12].Auto := 1, [0,12].Manual := 1, [0,12].OpenStatus := 1, [0,12].ZSOverride := 1, [0,12].FailState := 1, [0,12].EnableCfg := 1, [0,12].StatusWord := 2, [0,12].Status := 2, [0,12].OutputAddress := 44, [0,12].AlarmTimer.PRE := 2000, [0,12].AlarmTimerSP := 2, [0,12].AutoCloseTimer.ACC := 1072, [0,13].Tag := 'XV014', [0,13].Control := 1, [0,13].Auto := 1, [0,13].Manual := 1, [0,13].OpenStatus := 1, [0,13].ZSOverride := 1, [0,13].FailState := 1, [0,13].EnableCfg := 1, [0,13].StatusWord := 2, [0,13].Status := 2, [0,13].OutputAddress := 45, [0,13].AlarmTimer.PRE := 2000, [0,13].AlarmTimerSP := 2, [0,13].AutoCloseTimer.ACC := 1016, [0,14].Tag := 'XV015', [0,14].CloseStatus := 1, [0,14].ZSOverride := 1, [0,14].EnableCfg := 1, [0,14].StatusWord := 4, [0,14].Status := 4, [0,14].OutputAddress := 46, [0,14].AlarmTimer.PRE := 2000, [0,14].AlarmTimerSP := 2, [0,15].Tag := 'XV016', [0,15].Control := 1, [0,15].Auto := 1, [0,15].Manual := 1, [0,15].OpenStatus := 1, [0,15].ZSOverride := 1, [0,15].FailState := 1, [0,15].EnableCfg := 1, [0,15].StatusWord := 2, [0,15].Status := 2, [0,15].OutputAddress := 47, [0,15].AlarmTimer.PRE := 2000, [0,15].AlarmTimerSP := 2, [0,16].Tag := 'XV017', [0,16].CloseStatus := 1, [0,16].ZSOverride := 1, [0,16].EnableCfg := 1, [0,16].StatusWord := 4, [0,16].Status := 4, [0,16].OutputAddress := 48,
        [0,16].AlarmTimer.PRE := 2000, [0,16].AlarmTimerSP := 2, [0,17].Tag := 'XV018', [0,17].Control := 1, [0,17].Auto := 1, [0,17].Manual := 1, [0,17].OpenStatus := 1, [0,17].ZSOverride := 1, [0,17].FailState := 1, [0,17].EnableCfg := 1, [0,17].StatusWord := 2, [0,17].Status := 2, [0,17].OutputAddress := 49, [0,17].AlarmTimer.PRE := 2000, [0,17].AlarmTimerSP := 2, [0,17].AutoCloseTimer.ACC := 1594, [0,18].Tag := 'XV019', [0,18].CloseStatus := 1, [0,18].ZSOverride := 1, [0,18].EnableCfg := 1, [0,18].StatusWord := 4, [0,18].Status := 4, [0,18].OutputAddress := 50, [0,18].AlarmTimer.PRE := 2000, [0,18].AlarmTimerSP := 2, [0,18].AutoCloseTimer.ACC := 137, [0,19].Tag := 'XV020', [0,19].CloseStatus := 1, [0,19].ZSOverride := 1, [0,19].EnableCfg := 1, [0,19].StatusWord := 4, [0,19].Status := 4, [0,19].OutputAddress := 51, [0,19].AlarmTimer.PRE := 2000, [0,19].AlarmTimerSP := 2, [0,19].AutoCloseTimer.ACC := 1007, [0,20].Tag := 'XV021', [0,20].CloseStatus := 1, [0,20].ZSOverride := 1, [0,20].EnableCfg := 1, [0,20].StatusWord := 4, [0,20].Status := 4, [0,20].OutputAddress := 52, [0,20].AlarmTimer.PRE := 2000, [0,20].AlarmTimerSP := 2, [0,20].AutoCloseTimer.ACC := 1004, [0,21].Tag := 'XV022', [0,21].Control := 1, [0,21].Auto := 1, [0,21].Manual := 1, [0,21].OpenStatus := 1, [0,21].ZSOverride := 1, [0,21].FailState := 1, [0,21].EnableCfg := 1, [0,21].StatusWord := 2, [0,21].Status := 2, [0,21].OutputAddress := 53, [0,21].AlarmTimer.PRE := 2000, [0,21].AlarmTimerSP := 2, [0,22].Tag := 'XV023',
        [0,22].CloseStatus := 1, [0,22].ZSOverride := 1, [0,22].EnableCfg := 1, [0,22].StatusWord := 4, [0,22].Status := 4, [0,22].OutputAddress := 54, [0,22].AlarmTimer.PRE := 2000, [0,22].AlarmTimerSP := 2, [0,22].AutoCloseTimer.ACC := 131, [0,23].Tag := 'XV024', [0,23].CloseStatus := 1, [0,23].ZSOverride := 1, [0,23].EnableCfg := 1, [0,23].StatusWord := 4, [0,23].Status := 4, [0,23].OutputAddress := 55, [0,23].AlarmTimer.PRE := 2000, [0,23].AlarmTimerSP := 2, [0,23].AutoCloseTimer.ACC := 1003, [0,24].Tag := 'XV025', [0,24].CloseStatus := 1, [0,24].ZSOverride := 1, [0,24].EnableCfg := 1, [0,24].StatusWord := 4, [0,24].Status := 4, [0,24].OutputAddress := 56, [0,24].AlarmTimer.PRE := 2000, [0,24].AlarmTimerSP := 2, [0,24].AutoCloseTimer.ACC := 1002, [0,25].Tag := 'XV026', [0,25].CloseStatus := 1, [0,25].ZSOverride := 1, [0,25].EnableCfg := 1, [0,25].StatusWord := 4, [0,25].Status := 4, [0,25].OutputAddress := 57, [0,25].AlarmTimer.PRE := 2000, [0,25].AlarmTimerSP := 2, [0,25].AutoCloseTimer.ACC := 1002, [0,26].Tag := 'XV028', [0,26].CloseStatus := 1, [0,26].ZSOverride := 1, [0,26].EnableCfg := 1, [0,26].StatusWord := 4, [0,26].Status := 4, [0,26].OutputAddress := 58, [0,26].AlarmTimer.PRE := 2000, [0,26].AlarmTimerSP := 2, [0,26].AutoCloseTimer.ACC := 1002, [0,27].Tag := 'XV029', [0,27].CloseStatus := 1, [0,27].ZSOverride := 1, [0,27].EnableCfg := 1, [0,27].StatusWord := 4, [0,27].Status := 4, [0,27].OutputAddress := 59, [0,27].AlarmTimer.PRE := 2000, [0,27].AlarmTimerSP := 2, [0,28].Tag := 'XV030', [0,28].CloseStatus := 1,
        [0,28].ZSOverride := 1, [0,28].EnableCfg := 1, [0,28].StatusWord := 4, [0,28].Status := 4, [0,28].OutputAddress := 60, [0,28].AlarmTimer.PRE := 2000, [0,28].AlarmTimerSP := 2, [0,29].Tag := 'XV031', [0,29].Control := 1, [0,29].Auto := 1, [0,29].Manual := 1, [0,29].OpenStatus := 1, [0,29].ZSOverride := 1, [0,29].FailState := 1, [0,29].EnableCfg := 1, [0,29].StatusWord := 2, [0,29].Status := 2, [0,29].OutputAddress := 61, [0,29].AlarmTimer.PRE := 2000, [0,29].AlarmTimerSP := 2, [0,29].AutoCloseTimer.ACC := 1068, [0,30].Tag := 'XV033', [0,30].CloseStatus := 1, [0,30].ZSOverride := 1, [0,30].EnableCfg := 1, [0,30].StatusWord := 4, [0,30].Status := 4, [0,30].OutputAddress := 62, [0,30].AlarmTimer.PRE := 2000, [0,30].AlarmTimerSP := 2, [0,30].AutoCloseTimer.ACC := 1069, [0,31].Tag := 'XV034', [0,31].CloseStatus := 1, [0,31].ZSOverride := 1, [0,31].EnableCfg := 1, [0,31].StatusWord := 4, [0,31].Status := 4, [0,31].OutputAddress := 63, [0,31].AlarmTimer.PRE := 2000, [0,31].AlarmTimerSP := 2, [0,31].AutoCloseTimer.ACC := 131, [0,32].CloseStatus := 1, [0,32].PriorityCfg := 1, [0,32].ZSOpenAddress := 32, [0,32].OutputAddress := 68, [0,32].AlarmTimer.PRE := 2000, [0,32].AlarmTimerSP := 2, [0,32].AutoCloseTimer.ACC := 1059, [0,33].OpenStatus := 1, [0,33].PriorityCfg := 1, [0,33].FailState := 1, [0,33].ZSCloseAddress := 33, [0,33].OutputAddress := 69, [0,33].AlarmTimer.PRE := 2000, [0,33].AlarmTimerSP := 2, [0,33].AutoCloseTimer.ACC := 1123, [0,34].OpenStatus := 1, [0,34].PriorityCfg := 1, [0,34].FailState := 1, [0,34].ZSCloseAddress := 34,
        [0,34].OutputAddress := 70, [0,34].AlarmTimer.PRE := 2000, [0,34].AlarmTimerSP := 2, [0,34].AutoCloseTimer.ACC := 1095, [0,35].OpenStatus := 1, [0,35].PriorityCfg := 1, [0,35].FailState := 1, [0,35].ZSCloseAddress := 35, [0,35].OutputAddress := 71, [0,35].AlarmTimer.PRE := 2000, [0,35].AlarmTimerSP := 2, [0,35].AutoCloseTimer.ACC := 1127, [0,36].OpenStatus := 1, [0,36].PriorityCfg := 1, [0,36].FailState := 1, [0,36].ZSCloseAddress := 36, [0,36].OutputAddress := 72, [0,36].AlarmTimer.PRE := 2000, [0,36].AlarmTimerSP := 2, [0,36].AutoCloseTimer.ACC := 1004, [0,37].CloseStatus := 1, [0,37].PriorityCfg := 1, [0,37].ZSOpenAddress := 37, [0,37].OutputAddress := 73, [0,37].AlarmTimer.PRE := 2000, [0,37].AlarmTimerSP := 2, [0,37].AutoCloseTimer.ACC := 1121, [0,38].CloseStatus := 1, [0,38].Priority := 1, [0,38].PriorityCfg := 1, [0,38].ZSOpenAddress := 38, [0,38].OutputAddress := 40, [0,38].AlarmTimer.PRE := 2000, [0,38].AlarmTimerSP := 2, [0,38].AutoCloseTimer.ACC := 1135, [0,39].CloseStatus := 1, [0,39].Priority := 1, [0,39].PriorityCfg := 1, [0,39].ZSOpenAddress := 39, [0,39].OutputAddress := 41, [0,39].AlarmTimer.PRE := 2000, [0,39].AlarmTimerSP := 2, [0,39].AutoCloseTimer.ACC := 1121, [0,40].CloseStatus := 1, [0,40].Priority := 1, [0,40].PriorityCfg := 1, [0,40].ZSOpenAddress := 40, [0,40].OutputAddress := 42, [0,40].AlarmTimer.PRE := 2000, [0,40].AlarmTimerSP := 2, [0,40].AutoCloseTimer.ACC := 1112, [0,41].CloseStatus := 1, [0,41].Priority := 1, [0,41].PriorityCfg := 1, [0,41].ZSOpenAddress := 41, [0,41].OutputAddress := 43, [0,41].AlarmTimer.PRE := 2000, [0,41].AlarmTimerSP := 2, [0,42].CloseStatus := 1, [0,42].Priority := 1,
        [0,42].PriorityCfg := 1, [0,42].ZSOpenAddress := 42, [0,42].OutputAddress := 44, [0,42].AlarmTimer.PRE := 2000, [0,42].AlarmTimerSP := 2, [0,43].CloseStatus := 1, [0,43].Priority := 1, [0,43].PriorityCfg := 1, [0,43].ZSOpenAddress := 43, [0,43].OutputAddress := 52, [0,43].AlarmTimer.PRE := 2000, [0,43].AlarmTimerSP := 2, [0,44].CloseStatus := 1, [0,44].Priority := 1, [0,44].PriorityCfg := 1, [0,44].ZSOpenAddress := 44, [0,44].OutputAddress := 53, [0,44].AlarmTimer.PRE := 2000, [0,44].AlarmTimerSP := 2, [0,45].CloseStatus := 1, [0,45].Priority := 1, [0,45].PriorityCfg := 1, [0,45].ZSOpenAddress := 45, [0,45].OutputAddress := 54, [0,45].AlarmTimer.PRE := 2000, [0,45].AlarmTimerSP := 2, [0,46].CloseStatus := 1, [0,46].Priority := 1, [0,46].PriorityCfg := 1, [0,46].ZSOpenAddress := 46, [0,46].OutputAddress := 55, [0,46].AlarmTimer.PRE := 2000, [0,46].AlarmTimerSP := 2, [0,47].OpenStatus := 1, [0,47].Priority := 1, [0,47].PriorityCfg := 1, [0,47].FailState := 1, [0,47].ZSCloseAddress := 47, [0,47].OutputAddress := 45, [0,47].AlarmTimer.PRE := 2000, [0,47].AlarmTimerSP := 2, [0,48].FailState := 1, [0,48].ZSCloseAddress := 48, [0,48].OutputAddress := 80, [0,49].FailState := 1, [0,49].ZSCloseAddress := 49, [0,49].OutputAddress := 81, [0,50].FailState := 1, [0,50].ZSCloseAddress := 50, [0,50].OutputAddress := 82, [0,51].OpenStatus := 1, [0,51].FailState := 1, [0,51].ZSCloseAddress := 51, [0,51].OutputAddress := 83, [0,52].OpenStatus := 1, [0,52].FailState := 1, [0,52].ZSCloseAddress := 52, [0,52].OutputAddress := 84, [0,53].CloseStatus := 1, [0,53].FailState := 1,
        [0,53].ZSCloseAddress := 53, [0,53].OutputAddress := 85, [0,54].CloseStatus := 1, [0,54].FailState := 1, [0,54].ZSCloseAddress := 54, [0,54].OutputAddress := 86, [0,55].CloseStatus := 1, [0,55].FailState := 1, [0,55].ZSCloseAddress := 55, [0,55].OutputAddress := 87, [0,56].CloseStatus := 1, [0,58].CloseStatus := 1, [0,59].CloseStatus := 1, [1,0].Tag := 'XV001', [1,0].CloseStatus := 1, [1,0].ZSOverride := 1, [1,0].EnableCfg := 1, [1,0].StatusWord := 4, [1,0].Status := 4, [1,0].OutputAddress := 32, [1,0].AlarmTimer.PRE := 2000, [1,0].AlarmTimerSP := 2, [1,1].Tag := 'XV002', [1,1].CloseStatus := 1, [1,1].ZSOverride := 1, [1,1].EnableCfg := 1, [1,1].StatusWord := 4, [1,1].Status := 4, [1,1].OutputAddress := 33, [1,1].AlarmTimer.PRE := 2000, [1,1].AlarmTimerSP := 2, [1,1].AutoCloseTimer.ACC := 1103, [1,2].Tag := 'XV003', [1,2].CloseStatus := 1, [1,2].ZSOverride := 1, [1,2].EnableCfg := 1, [1,2].StatusWord := 4, [1,2].Status := 4, [1,2].OutputAddress := 34, [1,2].AlarmTimer.PRE := 2000, [1,2].AlarmTimerSP := 2, [1,2].AutoCloseTimer.ACC := 1032, [1,3].Tag := 'XV004', [1,3].CloseStatus := 1, [1,3].ZSOverride := 1, [1,3].EnableCfg := 1, [1,3].StatusWord := 4, [1,3].Status := 4, [1,3].OutputAddress := 35, [1,3].AlarmTimer.PRE := 2000, [1,3].AlarmTimerSP := 2, [1,3].AutoCloseTimer.ACC := 1115, [1,4].Tag := 'XV005', [1,4].CloseStatus := 1, [1,4].ZSOverride := 1, [1,4].EnableCfg := 1, [1,4].StatusWord := 4, [1,4].Status := 4, [1,4].OutputAddress := 36, [1,4].AlarmTimer.PRE := 2000,
        [1,4].AlarmTimerSP := 2, [1,4].AutoCloseTimer.ACC := 1104, [1,5].Tag := 'XV006', [1,5].CloseStatus := 1, [1,5].ZSOverride := 1, [1,5].EnableCfg := 1, [1,5].StatusWord := 4, [1,5].Status := 4, [1,5].OutputAddress := 37, [1,5].AlarmTimer.PRE := 2000, [1,5].AlarmTimerSP := 2, [1,5].AutoCloseTimer.ACC := 1104, [1,6].Tag := 'XV007', [1,6].CloseStatus := 1, [1,6].ZSOverride := 1, [1,6].EnableCfg := 1, [1,6].StatusWord := 4, [1,6].Status := 4, [1,6].OutputAddress := 38, [1,6].AlarmTimer.PRE := 2000, [1,6].AlarmTimerSP := 2, [1,6].AutoCloseTimer.ACC := 1104, [1,7].Tag := 'XV008', [1,7].CloseStatus := 1, [1,7].ZSOverride := 1, [1,7].EnableCfg := 1, [1,7].StatusWord := 4, [1,7].Status := 4, [1,7].OutputAddress := 39, [1,7].AlarmTimer.PRE := 2000, [1,7].AlarmTimerSP := 2, [1,7].AutoCloseTimer.ACC := 1104, [1,8].Tag := 'XV009', [1,8].CloseStatus := 1, [1,8].ZSOverride := 1, [1,8].EnableCfg := 1, [1,8].StatusWord := 4, [1,8].Status := 4, [1,8].OutputAddress := 40, [1,8].AlarmTimer.PRE := 2000, [1,8].AlarmTimerSP := 2, [1,8].AutoCloseTimer.ACC := 1104, [1,9].Tag := 'XV010', [1,9].CloseStatus := 1, [1,9].ZSOverride := 1, [1,9].EnableCfg := 1, [1,9].StatusWord := 4, [1,9].Status := 4, [1,9].OutputAddress := 41, [1,9].AlarmTimer.PRE := 2000, [1,9].AlarmTimerSP := 2, [1,9].AutoCloseTimer.ACC := 1105, [1,10].Tag := 'XV011', [1,10].CloseStatus := 1, [1,10].ZSOverride := 1, [1,10].EnableCfg := 1, [1,10].StatusWord := 4, [1,10].Status := 4, [1,10].OutputAddress := 42, [1,10].AlarmTimer.PRE := 2000,
        [1,10].AlarmTimerSP := 2, [1,10].AutoCloseTimer.ACC := 1104, [1,11].Tag := 'XV012', [1,11].Control := 1, [1,11].Auto := 1, [1,11].Manual := 1, [1,11].OpenStatus := 1, [1,11].ZSOverride := 1, [1,11].FailState := 1, [1,11].EnableCfg := 1, [1,11].StatusWord := 2, [1,11].Status := 2, [1,11].OutputAddress := 43, [1,11].AlarmTimer.PRE := 2000, [1,11].AlarmTimerSP := 2, [1,11].AutoCloseTimer.ACC := 1103, [1,12].Tag := 'XV013', [1,12].Control := 1, [1,12].Auto := 1, [1,12].Manual := 1, [1,12].OpenStatus := 1, [1,12].ZSOverride := 1, [1,12].FailState := 1, [1,12].EnableCfg := 1, [1,12].StatusWord := 2, [1,12].Status := 2, [1,12].OutputAddress := 44, [1,12].AlarmTimer.PRE := 2000, [1,12].AlarmTimerSP := 2, [1,12].AutoCloseTimer.ACC := 1072, [1,13].Tag := 'XV014', [1,13].Control := 1, [1,13].Auto := 1, [1,13].Manual := 1, [1,13].OpenStatus := 1, [1,13].ZSOverride := 1, [1,13].FailState := 1, [1,13].EnableCfg := 1, [1,13].StatusWord := 2, [1,13].Status := 2, [1,13].OutputAddress := 45, [1,13].AlarmTimer.PRE := 2000, [1,13].AlarmTimerSP := 2, [1,13].AutoCloseTimer.ACC := 1016, [1,14].Tag := 'XV015', [1,14].CloseStatus := 1, [1,14].ZSOverride := 1, [1,14].EnableCfg := 1, [1,14].StatusWord := 4, [1,14].Status := 4, [1,14].OutputAddress := 46, [1,14].AlarmTimer.PRE := 2000, [1,14].AlarmTimerSP := 2, [1,15].Tag := 'XV016', [1,15].Control := 1, [1,15].Auto := 1, [1,15].Manual := 1, [1,15].OpenStatus := 1, [1,15].ZSOverride := 1, [1,15].FailState := 1,
        [1,15].EnableCfg := 1, [1,15].StatusWord := 2, [1,15].Status := 2, [1,15].OutputAddress := 47, [1,15].AlarmTimer.PRE := 2000, [1,15].AlarmTimerSP := 2, [1,16].Tag := 'XV017', [1,16].CloseStatus := 1, [1,16].ZSOverride := 1, [1,16].EnableCfg := 1, [1,16].StatusWord := 4, [1,16].Status := 4, [1,16].OutputAddress := 48, [1,16].AlarmTimer.PRE := 2000, [1,16].AlarmTimerSP := 2, [1,17].Tag := 'XV018', [1,17].Control := 1, [1,17].Auto := 1, [1,17].Manual := 1, [1,17].OpenStatus := 1, [1,17].ZSOverride := 1, [1,17].FailState := 1, [1,17].EnableCfg := 1, [1,17].StatusWord := 2, [1,17].Status := 2, [1,17].OutputAddress := 49, [1,17].AlarmTimer.PRE := 2000, [1,17].AlarmTimerSP := 2, [1,17].AutoCloseTimer.ACC := 1594, [1,18].Tag := 'XV019', [1,18].CloseStatus := 1, [1,18].ZSOverride := 1, [1,18].EnableCfg := 1, [1,18].StatusWord := 4, [1,18].Status := 4, [1,18].OutputAddress := 50, [1,18].AlarmTimer.PRE := 2000, [1,18].AlarmTimerSP := 2, [1,18].AutoCloseTimer.ACC := 137, [1,19].Tag := 'XV020', [1,19].CloseStatus := 1, [1,19].ZSOverride := 1, [1,19].EnableCfg := 1, [1,19].StatusWord := 4, [1,19].Status := 4, [1,19].OutputAddress := 51, [1,19].AlarmTimer.PRE := 2000, [1,19].AlarmTimerSP := 2, [1,19].AutoCloseTimer.ACC := 1007, [1,20].Tag := 'XV021', [1,20].CloseStatus := 1, [1,20].ZSOverride := 1, [1,20].EnableCfg := 1, [1,20].StatusWord := 4, [1,20].Status := 4, [1,20].OutputAddress := 52, [1,20].AlarmTimer.PRE := 2000, [1,20].AlarmTimerSP := 2, [1,20].AutoCloseTimer.ACC := 1004, [1,21].Tag := 'XV022',
        [1,21].Control := 1, [1,21].Auto := 1, [1,21].Manual := 1, [1,21].OpenStatus := 1, [1,21].ZSOverride := 1, [1,21].FailState := 1, [1,21].EnableCfg := 1, [1,21].StatusWord := 2, [1,21].Status := 2, [1,21].OutputAddress := 53, [1,21].AlarmTimer.PRE := 2000, [1,21].AlarmTimerSP := 2, [1,22].Tag := 'XV023', [1,22].CloseStatus := 1, [1,22].ZSOverride := 1, [1,22].EnableCfg := 1, [1,22].StatusWord := 4, [1,22].Status := 4, [1,22].OutputAddress := 54, [1,22].AlarmTimer.PRE := 2000, [1,22].AlarmTimerSP := 2, [1,22].AutoCloseTimer.ACC := 131, [1,23].Tag := 'XV024', [1,23].CloseStatus := 1, [1,23].ZSOverride := 1, [1,23].EnableCfg := 1, [1,23].StatusWord := 4, [1,23].Status := 4, [1,23].OutputAddress := 55, [1,23].AlarmTimer.PRE := 2000, [1,23].AlarmTimerSP := 2, [1,23].AutoCloseTimer.ACC := 1003, [1,24].Tag := 'XV025', [1,24].CloseStatus := 1, [1,24].ZSOverride := 1, [1,24].EnableCfg := 1, [1,24].StatusWord := 4, [1,24].Status := 4, [1,24].OutputAddress := 56, [1,24].AlarmTimer.PRE := 2000, [1,24].AlarmTimerSP := 2, [1,24].AutoCloseTimer.ACC := 1002, [1,25].Tag := 'XV026', [1,25].CloseStatus := 1, [1,25].ZSOverride := 1, [1,25].EnableCfg := 1, [1,25].StatusWord := 4, [1,25].Status := 4, [1,25].OutputAddress := 57, [1,25].AlarmTimer.PRE := 2000, [1,25].AlarmTimerSP := 2, [1,25].AutoCloseTimer.ACC := 1002, [1,26].Tag := 'XV028', [1,26].CloseStatus := 1, [1,26].ZSOverride := 1, [1,26].EnableCfg := 1, [1,26].StatusWord := 4, [1,26].Status := 4, [1,26].OutputAddress := 58, [1,26].AlarmTimer.PRE := 2000,
        [1,26].AlarmTimerSP := 2, [1,26].AutoCloseTimer.ACC := 1002, [1,27].Tag := 'XV029', [1,27].CloseStatus := 1, [1,27].ZSOverride := 1, [1,27].EnableCfg := 1, [1,27].StatusWord := 4, [1,27].Status := 4, [1,27].OutputAddress := 59, [1,27].AlarmTimer.PRE := 2000, [1,27].AlarmTimerSP := 2, [1,28].Tag := 'XV030', [1,28].CloseStatus := 1, [1,28].ZSOverride := 1, [1,28].EnableCfg := 1, [1,28].StatusWord := 4, [1,28].Status := 4, [1,28].OutputAddress := 60, [1,28].AlarmTimer.PRE := 2000, [1,28].AlarmTimerSP := 2, [1,29].Tag := 'XV031', [1,29].Control := 1, [1,29].Auto := 1, [1,29].Manual := 1, [1,29].OpenStatus := 1, [1,29].ZSOverride := 1, [1,29].FailState := 1, [1,29].EnableCfg := 1, [1,29].StatusWord := 2, [1,29].Status := 2, [1,29].OutputAddress := 61, [1,29].AlarmTimer.PRE := 2000, [1,29].AlarmTimerSP := 2, [1,29].AutoCloseTimer.ACC := 1068, [1,30].Tag := 'XV033', [1,30].CloseStatus := 1, [1,30].ZSOverride := 1, [1,30].EnableCfg := 1, [1,30].StatusWord := 4, [1,30].Status := 4, [1,30].OutputAddress := 62, [1,30].AlarmTimer.PRE := 2000, [1,30].AlarmTimerSP := 2, [1,30].AutoCloseTimer.ACC := 1069, [1,31].Tag := 'XV034', [1,31].CloseStatus := 1, [1,31].ZSOverride := 1, [1,31].EnableCfg := 1, [1,31].StatusWord := 4, [1,31].Status := 4, [1,31].OutputAddress := 63, [1,31].AlarmTimer.PRE := 2000, [1,31].AlarmTimerSP := 2, [1,31].AutoCloseTimer.ACC := 131, [1,32].CloseStatus := 1, [1,32].PriorityCfg := 1, [1,32].ZSOpenAddress := 32, [1,32].OutputAddress := 68, [1,32].AlarmTimer.PRE := 2000, [1,32].AlarmTimerSP := 2,
        [1,32].AutoCloseTimer.ACC := 1059, [1,33].OpenStatus := 1, [1,33].PriorityCfg := 1, [1,33].FailState := 1, [1,33].ZSCloseAddress := 33, [1,33].OutputAddress := 69, [1,33].AlarmTimer.PRE := 2000, [1,33].AlarmTimerSP := 2, [1,33].AutoCloseTimer.ACC := 1123, [1,34].OpenStatus := 1, [1,34].PriorityCfg := 1, [1,34].FailState := 1, [1,34].ZSCloseAddress := 34, [1,34].OutputAddress := 70, [1,34].AlarmTimer.PRE := 2000, [1,34].AlarmTimerSP := 2, [1,34].AutoCloseTimer.ACC := 1095, [1,35].OpenStatus := 1, [1,35].PriorityCfg := 1, [1,35].FailState := 1, [1,35].ZSCloseAddress := 35, [1,35].OutputAddress := 71, [1,35].AlarmTimer.PRE := 2000, [1,35].AlarmTimerSP := 2, [1,35].AutoCloseTimer.ACC := 1127, [1,36].OpenStatus := 1, [1,36].PriorityCfg := 1, [1,36].FailState := 1, [1,36].ZSCloseAddress := 36, [1,36].OutputAddress := 72, [1,36].AlarmTimer.PRE := 2000, [1,36].AlarmTimerSP := 2, [1,36].AutoCloseTimer.ACC := 1004, [1,37].CloseStatus := 1, [1,37].PriorityCfg := 1, [1,37].ZSOpenAddress := 37, [1,37].OutputAddress := 73, [1,37].AlarmTimer.PRE := 2000, [1,37].AlarmTimerSP := 2, [1,37].AutoCloseTimer.ACC := 1121, [1,38].CloseStatus := 1, [1,38].Priority := 1, [1,38].PriorityCfg := 1, [1,38].ZSOpenAddress := 38, [1,38].OutputAddress := 40, [1,38].AlarmTimer.PRE := 2000, [1,38].AlarmTimerSP := 2, [1,38].AutoCloseTimer.ACC := 1135, [1,39].CloseStatus := 1, [1,39].Priority := 1, [1,39].PriorityCfg := 1, [1,39].ZSOpenAddress := 39, [1,39].OutputAddress := 41, [1,39].AlarmTimer.PRE := 2000, [1,39].AlarmTimerSP := 2, [1,39].AutoCloseTimer.ACC := 1121, [1,40].CloseStatus := 1, [1,40].Priority := 1, [1,40].PriorityCfg := 1, [1,40].ZSOpenAddress := 40,
        [1,40].OutputAddress := 42, [1,40].AlarmTimer.PRE := 2000, [1,40].AlarmTimerSP := 2, [1,40].AutoCloseTimer.ACC := 1112, [1,41].CloseStatus := 1, [1,41].Priority := 1, [1,41].PriorityCfg := 1, [1,41].ZSOpenAddress := 41, [1,41].OutputAddress := 43, [1,41].AlarmTimer.PRE := 2000, [1,41].AlarmTimerSP := 2, [1,42].CloseStatus := 1, [1,42].Priority := 1, [1,42].PriorityCfg := 1, [1,42].ZSOpenAddress := 42, [1,42].OutputAddress := 44, [1,42].AlarmTimer.PRE := 2000, [1,42].AlarmTimerSP := 2, [1,43].CloseStatus := 1, [1,43].Priority := 1, [1,43].PriorityCfg := 1, [1,43].ZSOpenAddress := 43, [1,43].OutputAddress := 52, [1,43].AlarmTimer.PRE := 2000, [1,43].AlarmTimerSP := 2, [1,44].CloseStatus := 1, [1,44].Priority := 1, [1,44].PriorityCfg := 1, [1,44].ZSOpenAddress := 44, [1,44].OutputAddress := 53, [1,44].AlarmTimer.PRE := 2000, [1,44].AlarmTimerSP := 2, [1,45].CloseStatus := 1, [1,45].Priority := 1, [1,45].PriorityCfg := 1, [1,45].ZSOpenAddress := 45, [1,45].OutputAddress := 54, [1,45].AlarmTimer.PRE := 2000, [1,45].AlarmTimerSP := 2, [1,46].CloseStatus := 1, [1,46].Priority := 1, [1,46].PriorityCfg := 1, [1,46].ZSOpenAddress := 46, [1,46].OutputAddress := 55, [1,46].AlarmTimer.PRE := 2000, [1,46].AlarmTimerSP := 2, [1,47].OpenStatus := 1, [1,47].Priority := 1, [1,47].PriorityCfg := 1, [1,47].FailState := 1, [1,47].ZSCloseAddress := 47, [1,47].OutputAddress := 45, [1,47].AlarmTimer.PRE := 2000, [1,47].AlarmTimerSP := 2, [1,48].FailState := 1, [1,48].ZSCloseAddress := 48, [1,48].OutputAddress := 80, [1,49].FailState := 1, [1,49].ZSCloseAddress := 49, [1,49].OutputAddress := 81,
        [1,50].FailState := 1, [1,50].ZSCloseAddress := 50, [1,50].OutputAddress := 82, [1,51].OpenStatus := 1, [1,51].FailState := 1, [1,51].ZSCloseAddress := 51, [1,51].OutputAddress := 83, [1,52].OpenStatus := 1, [1,52].FailState := 1, [1,52].ZSCloseAddress := 52, [1,52].OutputAddress := 84, [1,53].CloseStatus := 1, [1,53].FailState := 1, [1,53].ZSCloseAddress := 53, [1,53].OutputAddress := 85, [1,54].CloseStatus := 1, [1,54].FailState := 1, [1,54].ZSCloseAddress := 54, [1,54].OutputAddress := 86, [1,55].CloseStatus := 1, [1,55].FailState := 1, [1,55].ZSCloseAddress := 55, [1,55].OutputAddress := 87, [1,56].CloseStatus := 1, [1,58].CloseStatus := 1, [1,59].CloseStatus := 1, [2,0].Tag := 'XV001', [2,0].CloseStatus := 1, [2,0].ZSOverride := 1, [2,0].EnableCfg := 1, [2,0].StatusWord := 4, [2,0].Status := 4, [2,0].OutputAddress := 32, [2,0].AlarmTimer.PRE := 2000, [2,0].AlarmTimerSP := 2, [2,1].Tag := 'XV002', [2,1].CloseStatus := 1, [2,1].ZSOverride := 1, [2,1].EnableCfg := 1, [2,1].StatusWord := 4, [2,1].Status := 4, [2,1].OutputAddress := 33, [2,1].AlarmTimer.PRE := 2000, [2,1].AlarmTimerSP := 2, [2,1].AutoCloseTimer.ACC := 1103, [2,2].Tag := 'XV003', [2,2].CloseStatus := 1, [2,2].ZSOverride := 1, [2,2].EnableCfg := 1, [2,2].StatusWord := 4, [2,2].Status := 4, [2,2].OutputAddress := 34, [2,2].AlarmTimer.PRE := 2000, [2,2].AlarmTimerSP := 2, [2,2].AutoCloseTimer.ACC := 1032, [2,3].Tag := 'XV004', [2,3].CloseStatus := 1, [2,3].ZSOverride := 1, [2,3].EnableCfg := 1, [2,3].StatusWord := 4,
        [2,3].Status := 4, [2,3].OutputAddress := 35, [2,3].AlarmTimer.PRE := 2000, [2,3].AlarmTimerSP := 2, [2,3].AutoCloseTimer.ACC := 1115, [2,4].Tag := 'XV005', [2,4].CloseStatus := 1, [2,4].ZSOverride := 1, [2,4].EnableCfg := 1, [2,4].StatusWord := 4, [2,4].Status := 4, [2,4].OutputAddress := 36, [2,4].AlarmTimer.PRE := 2000, [2,4].AlarmTimerSP := 2, [2,4].AutoCloseTimer.ACC := 1104, [2,5].Tag := 'XV006', [2,5].CloseStatus := 1, [2,5].ZSOverride := 1, [2,5].EnableCfg := 1, [2,5].StatusWord := 4, [2,5].Status := 4, [2,5].OutputAddress := 37, [2,5].AlarmTimer.PRE := 2000, [2,5].AlarmTimerSP := 2, [2,5].AutoCloseTimer.ACC := 1104, [2,6].Tag := 'XV007', [2,6].CloseStatus := 1, [2,6].ZSOverride := 1, [2,6].EnableCfg := 1, [2,6].StatusWord := 4, [2,6].Status := 4, [2,6].OutputAddress := 38, [2,6].AlarmTimer.PRE := 2000, [2,6].AlarmTimerSP := 2, [2,6].AutoCloseTimer.ACC := 1104, [2,7].Tag := 'XV008', [2,7].CloseStatus := 1, [2,7].ZSOverride := 1, [2,7].EnableCfg := 1, [2,7].StatusWord := 4, [2,7].Status := 4, [2,7].OutputAddress := 39, [2,7].AlarmTimer.PRE := 2000, [2,7].AlarmTimerSP := 2, [2,7].AutoCloseTimer.ACC := 1104, [2,8].Tag := 'XV009', [2,8].CloseStatus := 1, [2,8].ZSOverride := 1, [2,8].EnableCfg := 1, [2,8].StatusWord := 4, [2,8].Status := 4, [2,8].OutputAddress := 40, [2,8].AlarmTimer.PRE := 2000, [2,8].AlarmTimerSP := 2, [2,8].AutoCloseTimer.ACC := 1104, [2,9].Tag := 'XV010', [2,9].CloseStatus := 1, [2,9].ZSOverride := 1, [2,9].EnableCfg := 1, [2,9].StatusWord := 4,
        [2,9].Status := 4, [2,9].OutputAddress := 41, [2,9].AlarmTimer.PRE := 2000, [2,9].AlarmTimerSP := 2, [2,9].AutoCloseTimer.ACC := 1105, [2,10].Tag := 'XV011', [2,10].CloseStatus := 1, [2,10].ZSOverride := 1, [2,10].EnableCfg := 1, [2,10].StatusWord := 4, [2,10].Status := 4, [2,10].OutputAddress := 42, [2,10].AlarmTimer.PRE := 2000, [2,10].AlarmTimerSP := 2, [2,10].AutoCloseTimer.ACC := 1104, [2,11].Tag := 'XV012', [2,11].Control := 1, [2,11].Auto := 1, [2,11].Manual := 1, [2,11].OpenStatus := 1, [2,11].ZSOverride := 1, [2,11].FailState := 1, [2,11].EnableCfg := 1, [2,11].StatusWord := 2, [2,11].Status := 2, [2,11].OutputAddress := 43, [2,11].AlarmTimer.PRE := 2000, [2,11].AlarmTimerSP := 2, [2,11].AutoCloseTimer.ACC := 1103, [2,12].Tag := 'XV013', [2,12].Control := 1, [2,12].Auto := 1, [2,12].Manual := 1, [2,12].OpenStatus := 1, [2,12].ZSOverride := 1, [2,12].FailState := 1, [2,12].EnableCfg := 1, [2,12].StatusWord := 2, [2,12].Status := 2, [2,12].OutputAddress := 44, [2,12].AlarmTimer.PRE := 2000, [2,12].AlarmTimerSP := 2, [2,12].AutoCloseTimer.ACC := 1072, [2,13].Tag := 'XV014', [2,13].Control := 1, [2,13].Auto := 1, [2,13].Manual := 1, [2,13].OpenStatus := 1, [2,13].ZSOverride := 1, [2,13].FailState := 1, [2,13].EnableCfg := 1, [2,13].StatusWord := 2, [2,13].Status := 2, [2,13].OutputAddress := 45, [2,13].AlarmTimer.PRE := 2000, [2,13].AlarmTimerSP := 2, [2,13].AutoCloseTimer.ACC := 1016, [2,14].Tag := 'XV015', [2,14].CloseStatus := 1, [2,14].ZSOverride := 1,
        [2,14].EnableCfg := 1, [2,14].StatusWord := 4, [2,14].Status := 4, [2,14].OutputAddress := 46, [2,14].AlarmTimer.PRE := 2000, [2,14].AlarmTimerSP := 2, [2,15].Tag := 'XV016', [2,15].Control := 1, [2,15].Auto := 1, [2,15].Manual := 1, [2,15].OpenStatus := 1, [2,15].ZSOverride := 1, [2,15].FailState := 1, [2,15].EnableCfg := 1, [2,15].StatusWord := 2, [2,15].Status := 2, [2,15].OutputAddress := 47, [2,15].AlarmTimer.PRE := 2000, [2,15].AlarmTimerSP := 2, [2,16].Tag := 'XV017', [2,16].CloseStatus := 1, [2,16].ZSOverride := 1, [2,16].EnableCfg := 1, [2,16].StatusWord := 4, [2,16].Status := 4, [2,16].OutputAddress := 48, [2,16].AlarmTimer.PRE := 2000, [2,16].AlarmTimerSP := 2, [2,17].Tag := 'XV018', [2,17].Control := 1, [2,17].Auto := 1, [2,17].Manual := 1, [2,17].OpenStatus := 1, [2,17].ZSOverride := 1, [2,17].FailState := 1, [2,17].EnableCfg := 1, [2,17].StatusWord := 2, [2,17].Status := 2, [2,17].OutputAddress := 49, [2,17].AlarmTimer.PRE := 2000, [2,17].AlarmTimerSP := 2, [2,17].AutoCloseTimer.ACC := 1594, [2,18].Tag := 'XV019', [2,18].CloseStatus := 1, [2,18].ZSOverride := 1, [2,18].EnableCfg := 1, [2,18].StatusWord := 4, [2,18].Status := 4, [2,18].OutputAddress := 50, [2,18].AlarmTimer.PRE := 2000, [2,18].AlarmTimerSP := 2, [2,18].AutoCloseTimer.ACC := 137, [2,19].Tag := 'XV020', [2,19].CloseStatus := 1, [2,19].ZSOverride := 1, [2,19].EnableCfg := 1, [2,19].StatusWord := 4, [2,19].Status := 4, [2,19].OutputAddress := 51, [2,19].AlarmTimer.PRE := 2000,
